{region 'Documentation'}
(*!
<summary>Neutral or held technical Error; task completion is reported separately.</summary>
*)
{endregion}
{attribute 'monitoring' := 'call'}
PROPERTY Result : E_Result //! Neutral or held technical Error; task completion is reported separately.
GET // PUBLIC
END_GET
END_PROPERTY

END_INTERFACE

// ---- Framework/Common/Interfaces/I_ResultAggregator.TcIO
{region 'Documentation'}
(*!
<summary>Contribution-only view of an owner-held result collection. Reset and result/counter access remain with the owner.</summary>
<description>
The owner resets and reads its concrete collection; a contribution hook only adds each owned result once. Contributions are immediate, not subscriptions, and no provider reference is retained. The owner limits a collection to 65535 contributions. Total includes neutral and Abort outcomes as well as Passed, Failed and Error; logging severity is a separate domain.
</description>
*)
{endregion}
INTERFACE I_ResultAggregator

{region 'Documentation'}
(*!
<summary>Adds one provider result immediately; a null provider contributes one Error. No provider reference is retained.</summary>
*)
{endregion}
METHOD AddProvider
VAR_INPUT
    Provider : I_ResultProvider; //! Result provider read immediately; zero contributes Error. No reference is retained.
END_VAR
END_METHOD

{region 'Documentation'}
(*!
<summary>Counts one contribution and combines Error &gt; Abort &gt; Failed &gt; Passed &gt; NotEvaluated.</summary>
*)
{endregion}
METHOD AddResult
VAR_INPUT
    Result : E_Result; //! Evaluation result to count as one contribution; severity is Error > Abort > Failed > Passed > NotEvaluated.
END_VAR
END_METHOD

END_INTERFACE

// ---- Framework/Common/Interfaces/I_ResultProvider.TcIO
{region 'Documentation'}
(*!
<summary>Read-only identity and result view; queries do not advance or modify the provider.</summary>
*)
{endregion}
INTERFACE I_ResultProvider

{region 'Documentation'}
(*!
<summary>Hierarchical identity supplied by the owning initialization path.</summary>
*)
{endregion}
{attribute 'monitoring' := 'variable'}
PROPERTY Name : STRING(GVL_Constants.NameLength) //! Hierarchical identity supplied by the owning initialization path.
GET // PUBLIC
END_GET
END_PROPERTY

{region 'Documentation'}
(*!
<summary>Current result by value; reading has no processing side effects.</summary>
*)
{endregion}
{attribute 'monitoring' := 'call'}
PROPERTY Result : E_Result //! Current result by value; reading has no processing side effects.
GET // PUBLIC
END_GET
END_PROPERTY

END_INTERFACE

// ---- Framework/EventBuffer/Interfaces/I_EventBuffer.TcIO
{region 'Documentation'}
(*!
<summary>Event storage initialization, administration, and value snapshots.</summary>
<description>
Bind one-based event storage and producer-owned status fields before administration. Keep them alive and stable and reinitialize after online change. The default service is single-task. Exactly one logical consumer acknowledges an epoch. External command handling and hierarchical reservation release belong to Run Control rather than this interface.
</description>
*)
{endregion}
INTERFACE I_EventBuffer

{region 'Documentation'}
(*!
<summary>Value snapshot of readable-range metadata.</summary>
*)
{endregion}
{attribute 'monitoring' := 'variable'}
PROPERTY FifoStatus : ST_FifoStatus //! Value snapshot of readable-range metadata.
GET // PUBLIC
END_GET
END_PROPERTY

{region 'Documentation'}
(*!
<summary>Bind one-based event storage and its producer-owned status fields for the service lifetime.</summary>
<description>
Establish an empty epoch; update the status fields internally after storage operations.

The default service requires lower bound 1 and physical length 3..32767; one ring position remains unused. Successful initialization clears the payload and begins a new empty epoch. Initialize owner reservation ledgers consistently; isolated reinitialization during execution is unsupported.
</description>
*)
{endregion}
METHOD Initialize : BOOL //! TRUE when storage is bound and usable; FALSE leaves the service uninitialized.
VAR_IN_OUT
    Buffer : ARRAY[*] OF ST_Event; //! Caller-owned event array, bound by address until reinitialization; keep storage alive and unchanged.
    FifoControl : ST_FifoStatus; //! Caller-owned FIFO status storage, retained and updated after buffer operations; must outlive the service.
    Status : ST_EventBufferStatus; //! Caller-owned event-sequence/loss snapshot, retained and updated by the service; must outlive it.
END_VAR
END_METHOD

{region 'Documentation'}
(*!
<summary>Release through the captured watermark; clear the caller&#x27;s field only if unchanged.</summary>
<description>
Use a current-epoch contiguous watermark after processing all preceding unread events. Zero is a no-op. Rejection or partial progress can still clear an unchanged request; inspect the actual DeletedSequenceId rather than treating command clearing as successful acknowledgement.
</description>
*)
{endregion}
METHOD ProcessDeleteRequest
VAR_IN_OUT
    SequenceId : UDINT; //! Inclusive deletion watermark; zero means no request. Cleared only if unchanged after processing.
END_VAR
END_METHOD

{region 'Documentation'}
(*!
<summary>Clear storage and epoch state while retaining a valid initialized binding.</summary>
<description>
A valid binding is required. The default service clears event storage, FIFO state, sequence, deletion watermark, loss count and aggregate reservations, retaining the binding. Owner-local accounting and external commands are handled by the Run Control integration path; they are not repaired here. Old-epoch acknowledgements become invalid.
</description>
*)
{endregion}
METHOD Reset
END_METHOD

{region 'Documentation'}
(*!
<summary>Value snapshot of sequence, deletion and loss status.</summary>
*)
{endregion}
{attribute 'monitoring' := 'variable'}
PROPERTY Status : ST_EventBufferStatus //! Value snapshot of sequence, deletion and loss status.
GET // PUBLIC
END_GET
END_PROPERTY

END_INTERFACE

// ---- Framework/EventBuffer/Interfaces/I_EventPublisher.TcIO
{region 'Documentation'}
(*!
<summary>PLC-side event publication and capacity view.</summary>
<description>
The default service is single-task and must be initialized with valid, stable storage before use. Publication copies the payload and assigns sequence/time; it does not consume an owner's reservation. Reservations are admission accounting, not storage or per-publication protection. Keep owner contributions consistent with the aggregate count and release them through their owner operations. Sequence exhaustion within an epoch is unsupported.
</description>
*)
{endregion}
INTERFACE I_EventPublisher

{region 'Documentation'}
(*!
<summary>Usable event positions, independent of occupancy and reservations; zero when invalid.</summary>
*)
{endregion}
{attribute 'monitoring' := 'call'}
PROPERTY Capacity : UINT //! Usable event positions, independent of occupancy and reservations; zero when invalid.
GET // PUBLIC
END_GET
END_PROPERTY

{region 'Documentation'}
(*!
<summary>Usable free event positions before reservations; zero when invalid.</summary>
*)
{endregion}
{attribute 'monitoring' := 'call'}
PROPERTY FreeEntryCount : UINT //! Usable free event positions before reservations; zero when invalid.
GET // PUBLIC
END_GET
END_PROPERTY

{region 'Documentation'}
(*!
<summary>Release only reservations, never events; FALSE changes neither count.</summary>
<description>
Requires an initialized valid binding, but no free capacity or valid FIFO indices.

The default service validates configuration and accounting even for a zero release. Free capacity and valid FIFO indices are not required. Destructive buffer reset clears the aggregate ledger, not stale owner-local contributions; use the coordinated owner release/reset path.
</description>
*)
{endregion}
METHOD FreeReservedSpace : BOOL //! TRUE after updating both reservation counts; FALSE leaves both unchanged.
VAR_INPUT
    EntryCount : UINT; //! Number of this owner's reserved entries to release; does not delete events.
END_VAR
VAR_IN_OUT
    OwnerReservedEntryCount : UINT; //! Owner's live reservation ledger; updated with the global count only on success, unchanged on rejection.
END_VAR
END_METHOD

{region 'Documentation'}
(*!
<summary>FIFO binding, configuration and indices are valid.</summary>
*)
{endregion}
{attribute 'monitoring' := 'call'}
PROPERTY IsValid : BOOL //! FIFO binding, configuration and indices are valid.
GET // PUBLIC
END_GET
END_PROPERTY

{region 'Documentation'}
(*!
<summary>Lost event count for producer diagnostics and aggregation.</summary>
*)
{endregion}
{attribute 'monitoring' := 'call'}
PROPERTY LostEventCount : UINT //! Lost event count for producer diagnostics and aggregation.
GET // PUBLIC
END_GET
END_PROPERTY

{region 'Documentation'}
(*!
<summary>Publish a value copy with producer-assigned SequenceId and UTC Timestamp.</summary>
<description>
Positive slot on success, zero when full, negative E_EventPublishResult on error.

The return describes the requested event. The default service may also attempt a capacity diagnostic after a successful insertion. That attempt can consume capacity or increase LostEventCount without changing the primary return. Publishing does not decrement an owner's reservation. Sequence numbers may be assigned before insertion succeeds; a nonzero loss count means an incomplete log.
</description>
*)
{endregion}
METHOD PublishEvent : INT //! Positive physical slot on success, zero when full, negative E_EventPublishResult on error.
VAR_INPUT
    Event : ST_Event; //! Event payload copied into the buffer; SequenceId and Timestamp are assigned by the publisher.
END_VAR
END_METHOD

{region 'Documentation'}
(*!
<summary>Aggregate producer reservations; not published externally.</summary>
*)
{endregion}
{attribute 'monitoring' := 'call'}
PROPERTY ReservedEntryCount : UINT //! Aggregate producer reservations; not published externally.
GET // PUBLIC
END_GET
END_PROPERTY

{region 'Documentation'}
(*!
<summary>Reserve additional event positions plus shared headroom; FALSE changes neither count.</summary>
<description>
Requires valid initialized configuration and a consistent owner contribution; positive requests also require valid indices.

For the default service, positive requests require free capacity for the updated aggregate count plus shared headroom. A zero request checks configuration and owner contribution but bypasses index and capacity checks. Both ledgers change together on success; no event is created. Keep the owner ledger unchanged by unrelated code.
</description>
*)
{endregion}
METHOD ReserveSpace : BOOL //! TRUE after updating both reservation counts; FALSE leaves both unchanged.
VAR_INPUT
    EntryCount : UINT; //! Additional number of event entries to reserve for this owner.
    HeadroomEntryCount : UINT; //! Shared free entries checked for positive requests; not added to the owner's reservation.
END_VAR
VAR_IN_OUT
    OwnerReservedEntryCount : UINT; //! Owner's live reservation ledger; updated with the global count only on success, unchanged on rejection.
END_VAR
END_METHOD

END_INTERFACE

// ---- Framework/Preparation/Interfaces/I_Preparation.TcIO
{region 'Documentation'}
(*!
<summary>Read-only Preparation view; querying does not execute resource actions.</summary>
<description>
This interface exposes only the last reported Status by value. The owner calls the concrete Preparation cyclically with Enable and its resource-specific bindings; the interface provides no generic activation, initialization or reset operation.
</description>
*)
{endregion}
INTERFACE I_Preparation

{region 'Documentation'}
(*!
<summary>Current Preparation status by value; querying does not execute resource actions.</summary>
*)
{endregion}
PROPERTY Status : ST_PreparationStatus //! Current Preparation status by value; querying does not execute resource actions.
GET // PUBLIC
END_GET
END_PROPERTY

END_INTERFACE

// ---- Framework/RunControl/Interfaces/I_RunControl.TcIO
{region 'Documentation'}
(*!
<summary>Run Control request and status view; the execution owner calls the concrete FB cyclically.</summary>
<description>
Request methods record same-task intent; they do not execute the lifecycle synchronously. Repeated requests coalesce and regular processing applies Reset over Abort over Start. Status is a stored value snapshot. Name and Result are inherited from I_ResultProvider. The concrete owner must still be called cyclically, including after completion.
</description>
*)
{endregion}
INTERFACE I_RunControl EXTENDS I_ResultProvider

{region 'Documentation'}
(*!
<summary>Records an abort request for regular lifecycle processing.</summary>
*)
{endregion}
METHOD RequestAbort
END_METHOD

{region 'Documentation'}
(*!
<summary>Records a reset request for regular lifecycle processing.</summary>
*)
{endregion}
METHOD RequestReset
END_METHOD

{region 'Documentation'}
(*!
<summary>Records a start request for regular lifecycle processing.</summary>
*)
{endregion}
METHOD RequestStart
END_METHOD

{region 'Documentation'}
(*!
<summary>Current owner status snapshot; reading does not execute lifecycle processing.</summary>
*)
{endregion}
PROPERTY Status : ST_RunControlStatus //! Current owner status snapshot; reading does not execute lifecycle processing.
GET // PUBLIC
END_GET
END_PROPERTY

END_INTERFACE

// ---- Framework/TestCases/Interfaces/I_TestCase.TcIO
{region 'Documentation'}
(*!
<summary>Typed owner status with the shared child orchestration view.</summary>
<description>
Adds only the typed Status snapshot to I_Orchestratable. Lifecycle requests, readiness/state, initialization, reservation operations, execution slot and inherited identity/result belong to that shared child view. Requests do not execute the concrete FB. The owning Suite calls the concrete instance cyclically; status reads do not refresh it.
</description>
*)
{endregion}
INTERFACE I_TestCase EXTENDS I_Orchestratable

{region 'Documentation'}
(*!
<summary>Return the latest typed Test Case status by value without executing lifecycle, Preparation or Assertion work.</summary>
*)
{endregion}
PROPERTY Status : ST_TestCaseStatus //! Return the latest typed Test Case status by value without executing lifecycle, Preparation or Assertion work.
GET // PUBLIC
END_GET
END_PROPERTY

END_INTERFACE

// ---- Framework/TestSuites/Interfaces/I_TestSuite.TcIO
{region 'Documentation'}
(*!
<summary>Typed owner status with the shared child orchestration view.</summary>
<description>
Adds only typed Status to I_Orchestratable; shared requests, readiness/state, initialization, reservation operations, slot and inherited identity/result remain in that view. The owner invokes the concrete FB cyclically; interface requests and getters do not execute it. Production composition and the explicitly childless mock have different internal responsibilities.
</description>
*)
{endregion}
INTERFACE I_TestSuite EXTENDS I_Orchestratable

{region 'Documentation'}
(*!
<summary>Current owner status snapshot; reading does not execute lifecycle processing.</summary>
*)
{endregion}
PROPERTY Status : ST_TestSuiteStatus //! Current owner status snapshot; reading does not execute lifecycle processing.
GET // PUBLIC
END_GET
END_PROPERTY

END_INTERFACE

// ---- Runtime/MAIN.TcPOU
{region 'Documentation'}
(*!
<summary>Initializes the selftest hierarchy on the first task cycle and executes its command adapter and root.</summary>
<description>
Assign MAIN once to the single cyclic task that owns the hierarchy. A nonpositive current task
index skips all work. On FirstCycle, clear old commands through the adapter, initialize the
actual Event Stream storage/status, then initialize the SelfTests root with that same buffer service.
The library's default publisher must refer to the matching service before configuration diagnostics.

Normal processing calls the command adapter before the concrete root on every valid task call,
including after initialization failure or lifecycle completion. The stored initialization outcomes
are diagnostic values, not cyclic execution gates; failed owner setup prevents normal child work
inside the base. There is no automatic cyclic initialization retry or automatic Start of tests.

Successful root initialization queues its initial lifecycle Reset; readiness is established over
subsequent cycles. Rebuilding setup requires configuration reactivation or PLC Cold Reset and the
coordinated first-cycle path. Normal Stop/Start and lifecycle Reset do not rebuild configuration.
This executable selftest composition is outside the packaged library and consumer API reference.
</description>
*)
{endregion}
PROGRAM MAIN
VAR
    {attribute 'TcNoSymbol'}
    FRunControl : RunControl; //! Statically owned selftest root; invoked once after command intake on every valid task call.
    {attribute 'TcNoSymbol'}
    FCommandAdapter : RunControlCommandAdapter; //! Owner-local command sampler; initialized before the Event Buffer and called before the root.
    {attribute 'TcNoSymbol'}
    FEventBufferInitialized : BOOL; //! Last first-cycle Event Buffer initialization outcome; diagnostic only, not a cyclic call gate.
    {attribute 'TcNoSymbol'}
    FFrameworkInitialized : BOOL; //! Last first-cycle hierarchy initialization outcome; TRUE does not yet imply Idle or Ready.
END_VAR
VAR_TEMP
    TaskIndex : DINT; //! Current cyclic PLC task index; nonpositive values skip initialization and execution.
END_VAR

TaskIndex := Tc2_System.GETCURTASKINDEXEX();
IF TaskIndex <= 0 THEN
    RETURN;
END_IF;

IF TwinCAT_SystemInfoVarList._TaskInfo[TaskIndex].FirstCycle THEN
    FCommandAdapter.Initialize(ControlData := GVL_UnitTest.RunControl.ControlData);

    FEventBufferInitialized := GVL_EventBuffer.Instance.Initialize(Buffer := GVL_UnitTest.EventStream.Buffer,
        FifoControl := GVL_UnitTest.EventStream.FifoControl,
        Status := GVL_UnitTest.EventStream.Status);

    FFrameworkInitialized := FRunControl.Initialize(Name := 'SelfTests',
        EventBuffer := GVL_EventBuffer.Instance);
END_IF;

FCommandAdapter(RunControl := FRunControl,
    Commands := GVL_UnitTest.RunControl.ControlData.Cmd);
FRunControl(ControlData := GVL_UnitTest.RunControl.ControlData);

END_PROGRAM

// ---- SelfTests/RunControl/RunControl.TcPOU
{region 'Documentation'}
(*!
<summary>Composes the selftest Suites and forwards the external communication storage to the root base.</summary>
*)
{endregion}
FUNCTION_BLOCK RunControl EXTENDS RunControlBase
VAR
    FSmoke : TestSuite_Smoke;
    FPreparation : TestSuite_Preparation;
    FTestCaseLifecycle : TestSuite_TestCaseLifecycle;
    FOrchestratorTests : TestSuite_Orchestrator;
    FSerialOrchestration : TestSuite_SerialOrchestration;
    FParallelOrchestration : TestSuite_ParallelOrchestration;
    FParallelSlotsOrchestration : TestSuite_ParallelSlotsOrchestration;
    FSuiteBuilderTests : TestSuite_TestSuiteConfigurationBuilder;
    FRunControlBuilderTests : TestSuite_RunControlConfigurationBuilder;
    FTestSuites : ARRAY[1..SuiteCapacity] OF I_TestSuite;
    FTestSuiteLifecycle : TestSuite_TestSuiteLifecycle;
    FRunControlLifecycle : TestSuite_RunControlLifecycle;
    FCommandAdapter : TestSuite_CommandAdapter;
    FEventDelivery : TestSuite_EventDelivery;
    FEventReservation : TestSuite_EventReservation;
    FEventBufferReset : TestSuite_EventBufferReset;
    FAssertionLifecycle : TestSuite_AssertionLifecycle;
    FAssertionComparisons : TestSuite_AssertionComparisons;
    FAssertionFloatingPoint : TestSuite_AssertionFloatingPoint;
    FAssertionObservation : TestSuite_AssertionObservation;
    FAssertionText : TestSuite_AssertionText;
    FAssertionArrays : TestSuite_AssertionArrays;
    FAssertionVariants : TestSuite_AssertionVariants;
END_VAR
VAR CONSTANT
    SuiteCapacity : UINT := 22;
END_VAR

SUPER^(ControlData := ControlData);

{region 'Documentation'}
(*!
<summary>Initializes and registers the selftest Suites serially. Root and Suite Reset timeouts allow 15 seconds for event-consumer backpressure.</summary>
*)
{endregion}
METHOD PROTECTED Configure
VAR_IN_OUT
    // SA0167: Borrowed builder; VAR_IN_OUT creates no temporary instance.
    {attribute 'analysis' := '-167'}
    Builder : RunControlConfigurationBuilder; //! Borrowed owner configuration builder used only during this Configure call; register this owner's concrete children.
END_VAR
VAR
    SuiteConfig : ST_TestSuiteConfig;
END_VAR
FConfig.Timeout := T#60s;
FConfig.ResetTimeout := T#15s;
SuiteConfig.ResetTimeout := T#15s;

Builder.Initialize(Mode := E_OrchestrationMode.Serial,
    TestSuites := FTestSuites);

FSmoke.Initialize(Parent := THIS^,
    SuiteName := 'Smoke',
    Config := SuiteConfig);
Builder.Register(TestSuite := FSmoke);

FPreparation.Initialize(Parent := THIS^,
    SuiteName := 'Preparation',
    Config := SuiteConfig);
Builder.Register(TestSuite := FPreparation);

FTestCaseLifecycle.Initialize(Parent := THIS^,
    SuiteName := 'TestCaseLifecycle',
    Config := SuiteConfig);
Builder.Register(TestSuite := FTestCaseLifecycle);

FOrchestratorTests.Initialize(Parent := THIS^,
    SuiteName := 'Orchestrator',
    Config := SuiteConfig);
Builder.Register(TestSuite := FOrchestratorTests);

FSerialOrchestration.Initialize(Parent := THIS^,
    SuiteName := 'SerialOrchestration',
    Config := SuiteConfig);
Builder.Register(TestSuite := FSerialOrchestration);

FParallelOrchestration.Initialize(Parent := THIS^,
    SuiteName := 'ParallelOrchestration',
    Config := SuiteConfig);
Builder.Register(TestSuite := FParallelOrchestration);

FParallelSlotsOrchestration.Initialize(Parent := THIS^,
    SuiteName := 'ParallelSlotsOrchestration',
    Config := SuiteConfig);
Builder.Register(TestSuite := FParallelSlotsOrchestration);

FSuiteBuilderTests.Initialize(Parent := THIS^,
    SuiteName := 'SuiteBuilder',
    Config := SuiteConfig);
Builder.Register(TestSuite := FSuiteBuilderTests);

FRunControlBuilderTests.Initialize(Parent := THIS^,
    SuiteName := 'RunControlBuilder',
    Config := SuiteConfig);
Builder.Register(TestSuite := FRunControlBuilderTests);

FTestSuiteLifecycle.BindSubjectParent(Parent := THIS^);
FTestSuiteLifecycle.Initialize(Parent := THIS^,
    SuiteName := 'TestSuiteLifecycle',
    Config := SuiteConfig);
Builder.Register(TestSuite := FTestSuiteLifecycle);

FRunControlLifecycle.Initialize(Parent := THIS^,
    SuiteName := 'RunControlLifecycle',
    Config := SuiteConfig);
Builder.Register(TestSuite := FRunControlLifecycle);

FCommandAdapter.Initialize(Parent := THIS^,
    SuiteName := 'CommandAdapter',
    Config := SuiteConfig);
Builder.Register(TestSuite := FCommandAdapter);

FEventDelivery.Initialize(Parent := THIS^,
    SuiteName := 'EventDelivery',
    Config := SuiteConfig);
Builder.Register(TestSuite := FEventDelivery);

FEventReservation.BindSubjectParent(Parent := THIS^);
FEventReservation.Initialize(Parent := THIS^,
    SuiteName := 'EventReservation',
    Config := SuiteConfig);
Builder.Register(TestSuite := FEventReservation);

FEventBufferReset.Initialize(Parent := THIS^,
    SuiteName := 'EventBufferReset',
    Config := SuiteConfig);
Builder.Register(TestSuite := FEventBufferReset);

FAssertionLifecycle.Initialize(Parent := THIS^,
    SuiteName := 'AssertionLifecycle',
    Config := SuiteConfig);
Builder.Register(TestSuite := FAssertionLifecycle);

FAssertionComparisons.Initialize(Parent := THIS^,
    SuiteName := 'AssertionComparisons',
    Config := SuiteConfig);
Builder.Register(TestSuite := FAssertionComparisons);

FAssertionFloatingPoint.Initialize(Parent := THIS^,
    SuiteName := 'AssertionFloatingPoint',
    Config := SuiteConfig);
Builder.Register(TestSuite := FAssertionFloatingPoint);

FAssertionObservation.Initialize(Parent := THIS^,
    SuiteName := 'AssertionObservation',
    Config := SuiteConfig);
Builder.Register(TestSuite := FAssertionObservation);

FAssertionText.Initialize(Parent := THIS^,
    SuiteName := 'AssertionText',
    Config := SuiteConfig);
Builder.Register(TestSuite := FAssertionText);

FAssertionArrays.Initialize(Parent := THIS^,
    SuiteName := 'AssertionArrays',
    Config := SuiteConfig);
Builder.Register(TestSuite := FAssertionArrays);

FAssertionVariants.Initialize(Parent := THIS^,
    SuiteName := 'AssertionVariants',
    Config := SuiteConfig);
Builder.Register(TestSuite := FAssertionVariants);
END_METHOD

{region 'Documentation'}
(*!
<summary>Returns the registered Suite from the same array used during configuration.</summary>
*)
{endregion}
METHOD PUBLIC GetTestSuite : I_TestSuite //! Typed Suite interface at the original array index; zero when no entry is available.
VAR_INPUT
    Index : DINT; //! Original occupied child-array index, rather than an ordinal position.
END_VAR
GetTestSuite := 0;
IF (ChildCount = 0) OR (Index < ChildArrayLowerBound)
    OR (DINT_TO_LINT(Index) >= DINT_TO_LINT(ChildArrayLowerBound) + UINT_TO_LINT(ChildCount)) THEN
    RETURN;
END_IF;

GetTestSuite := FTestSuites[Index];
END_METHOD

{region 'Documentation'}
(*!
<summary>Calls each owned Suite once per initialized root cycle, including completion.</summary>
*)
{endregion}
METHOD PROTECTED ProcessTestSuites
FSmoke();
FPreparation();
FTestCaseLifecycle();
FOrchestratorTests();
FSerialOrchestration();
FParallelOrchestration();
FParallelSlotsOrchestration();
FSuiteBuilderTests();
FRunControlBuilderTests();

FTestSuiteLifecycle();
FRunControlLifecycle();

FCommandAdapter();

FEventDelivery();

FEventReservation();
FEventBufferReset();
FAssertionLifecycle();
FAssertionComparisons();
FAssertionFloatingPoint();
FAssertionObservation();

FAssertionText();

FAssertionArrays();
FAssertionVariants();
END_METHOD

END_FUNCTION_BLOCK

// ---- Framework/RunControl/POU/RunControlBase.TcPOU
{region 'Documentation'}
(*!
<summary>Root lifecycle and orchestration of the application's static Suite collection.</summary>
<description>
The PLC program initializes the Event Buffer and publisher before Initialize. Implement
Configure, GetTestSuite and ProcessTestSuites; forward ControlData to SUPER^() once per task
cycle.

Run the external command adapter before this FB. Buffer commands are handled first; only Name
and Status are projected after lifecycle processing. CompletionDelay belongs to this root, not to
its Orchestrator.

Continue cyclic calls after Completed so descendants can finish outstanding work and status
can refresh. This does not reopen the finalized root result.

In Completing, Result and Aggregation are published once before CompletionDelay elapses. The
final transition occurs on a later call even for zero delay. Invalid delay timing emits a diagnostic
and completes without changing published results.
</description>
*)
{endregion}
FUNCTION_BLOCK ABSTRACT RunControlBase IMPLEMENTS I_RunControl, I_OrchestratableCollection
VAR_IN_OUT
    ControlData : ST_RunControl; //! External communication storage; BufferCmd is processed first, Name and Status are projected last.
END_VAR
VAR
    /// Instance binding; derived test adapters may assign it before first use.
    FEventPublisher : I_EventPublisher;
    FName : STRING(GVL_Constants.NameLength);
    FResourceName : STRING(GVL_Constants.ResourceNameLength);
    FConfig : ST_RunConfig;
    FEventBuffer : I_EventBuffer;
    FCollectionConfiguration : ST_TestSuiteCollectionConfig;
    FOrchestrator : I_Orchestrator;
    FDefaultOrchestrator : Orchestrator;
    FInitialized : BOOL;
    FHasTimeout : BOOL;
    FHasResetTimeout : BOOL;
    FHasAbortTimeout : BOOL;
    FCheckingInitialization : BOOL;
    FConfigError : BOOL;
    FStatus : ST_RunControlStatus;
    FResult : E_Result := E_Result.NotEvaluated;
    FState : E_State := E_State.Uninitialized;
    FMethodRequests : ST_Command;
    FExecutionTimer : Stopwatch;
    FStateTimer : Stopwatch;
    FAggregator : ResultAggregator;
    FTestSuiteCountInactive : UINT;
    FTestSuiteCountIdle : UINT;
    FTestSuiteCountRunning : UINT;
    FTestSuiteCountCompleted : UINT;
    FTestSuiteCountError : UINT;
    FCollectionValid : BOOL;
    FChildrenError : BOOL;
    FChildrenAborted : BOOL;
    FChildrenCompleted : BOOL;
    FChildrenAbortFinished : BOOL;
    FFinalizationPublished : BOOL;
END_VAR
VAR_TEMP
    Requests : ST_Command;
    OrchestratorTask : E_OrchestratorTask;
END_VAR

ProcessBufferCommands(Commands := ControlData.BufferCmd);
ProcessRequests(InputRequests := FMethodRequests, Requests => Requests);

FExecutionTimer.Update();
FStateTimer.Update();

Sequencer(Requests := Requests);

IF IsInitialized THEN
    OrchestratorTask := MapOrchestratorTask(State := FState,
        CurrentTask := FOrchestrator.CurrentTask);
    FOrchestrator.Execute(Task := OrchestratorTask);

    ProcessTestSuites();
    AggregateResults();
END_IF;

UpdateResult();
UpdateStatus();
EmitFinalizationEvents();

ControlData.Name := FName;
ControlData.Status := FStatus;

{region 'Documentation'}
(*!
<summary>Aggregates results and execution counters after child calls; refreshes observations from the same snapshots.</summary>
*)
{endregion}
METHOD PRIVATE AggregateResults
VAR
    Count : UINT;
    FirstIndex : DINT;
    LastIndex : DINT;
    Index : LINT;
    ChildStatus : ST_TestSuiteStatus;
    ChildResult : E_Result;
END_VAR
Count := ChildCount;
FTestSuiteCountInactive := 0;
FTestSuiteCountIdle := 0;
FTestSuiteCountRunning := 0;
FTestSuiteCountCompleted := 0;
FTestSuiteCountError := 0;
FAggregator.Reset();
FCollectionValid := FALSE;
FChildrenCompleted := FALSE;
FChildrenAbortFinished := FALSE;
FChildrenError := FALSE;
FChildrenAborted := FALSE;

IF NOT FInitialized OR (Count = 0) THEN
    RETURN;
END_IF;
FirstIndex := ChildArrayLowerBound;
LastIndex := ChildArrayUpperBound;
IF DINT_TO_LINT(LastIndex) - DINT_TO_LINT(FirstIndex) + 1 < UINT_TO_LINT(Count) THEN
    RETURN;
END_IF;

FCollectionValid := TRUE;
FChildrenCompleted := TRUE;
FChildrenAbortFinished := TRUE;
FOR Index := DINT_TO_LINT(FirstIndex) TO DINT_TO_LINT(FirstIndex) + UINT_TO_LINT(Count) - 1 DO
    IF NOT ObserveTestSuite(Child := GetTestSuite(Index := LINT_TO_DINT(Index)),
        ChildStatus => ChildStatus) THEN
        FTestSuiteCountError := FTestSuiteCountError + 1;
        FAggregator.AddResult(Result := E_Result.Error);
        CONTINUE;
    END_IF;

    ChildResult := ChildStatus.Execution.Result;
    CASE ChildResult OF
        E_Result.NotEvaluated, E_Result.Passed, E_Result.Failed, E_Result.Abort, E_Result.Error:
            FAggregator.AddResult(Result := ChildResult);
    ELSE
        ChildResult := E_Result.Error;
        FAggregator.AddResult(Result := ChildResult);
    END_CASE;

    CASE ChildStatus.Execution.ExecutionStatus OF
        E_ExecutionStatus.Inactive:
            FTestSuiteCountInactive := FTestSuiteCountInactive + 1;
        E_ExecutionStatus.Idle:
            FTestSuiteCountIdle := FTestSuiteCountIdle + 1;
        E_ExecutionStatus.Running:
            FTestSuiteCountRunning := FTestSuiteCountRunning + 1;
        E_ExecutionStatus.Completed:
            FTestSuiteCountCompleted := FTestSuiteCountCompleted + 1;
    ELSE
        // Transitional execution states have no dedicated counter in the status contract.
    END_CASE;
    IF (ChildStatus.Execution.ExecutionStatus = E_ExecutionStatus.Error) OR (ChildResult = E_Result.Error) THEN
        FTestSuiteCountError := FTestSuiteCountError + 1;
    END_IF;

END_FOR;
END_METHOD

{region 'Documentation'}
(*!
<summary>Applies permitted owner transitions; rejects others with state-dependent diagnostics and Error escalation while leaving FState unchanged.</summary>
*)
{endregion}
METHOD PRIVATE ChangeState
VAR_INPUT
    NewState : E_State; //! Requested owner lifecycle destination; identical state is a no-op and rejected transitions do not change FState.
END_VAR
IF NewState = FState THEN
    RETURN;
END_IF;
IF NOT IsStateTransitionAllowed(NewState := NewState) THEN
    CASE FState OF
        E_State.Uninitialized:
            RETURN;

        E_State.Completing, E_State.Completed:
            PublishEvent(Event := CreateInvalidStateTransitionEvent(OwnerScope := E_OwnerScope.RunControl,
                Name := FName,
                ResourceName := FResourceName,
                StateOld := FState,
                StateNew := NewState));
    ELSE
        IF FResult <> E_Result.Error THEN
            PublishEvent(Event := CreateInvalidStateTransitionEvent(OwnerScope := E_OwnerScope.RunControl,
                Name := FName,
                ResourceName := FResourceName,
                StateOld := FState,
                StateNew := NewState));
        END_IF;
        FResult := E_Result.Error;
    END_CASE;
    RETURN;
END_IF;

CASE NewState OF
    E_State.Uninitialized:
        FExecutionTimer.Reset();
        FStateTimer.Start();
        FResult := E_Result.NotEvaluated;
    E_State.Reset:
        FHasTimeout := FALSE;
        FHasResetTimeout := FALSE;
        FHasAbortTimeout := FALSE;
        FFinalizationPublished := FALSE;
        FAggregator.Reset();
        IF (FState = E_State.Starting) OR (FState = E_State.Running) OR (FState = E_State.Completing)
            OR (FState = E_State.Aborting) OR (FState = E_State.AbortingFromError) THEN
            PublishEvent(Event := CreateResetWarningEvent(OwnerScope := E_OwnerScope.RunControl,
                Name := FName,
                ResourceName := FResourceName,
                State := FState));
        END_IF;
        FExecutionTimer.Reset();
        FStateTimer.Start();
        FResult := E_Result.NotEvaluated;
    E_State.Idle:
        FStateTimer.Start();
    E_State.Starting:
        FStateTimer.Start();
        FExecutionTimer.Start();
    E_State.Running:
        FStateTimer.Start();
    E_State.Completing:
        FExecutionTimer.Stop();
        FStateTimer.Start();
    E_State.Completed:
        FStateTimer.Start();
    E_State.Aborting:
        FExecutionTimer.Stop();
        FStateTimer.Start();
        IF FResult <> E_Result.Error THEN
            FResult := E_Result.Abort;
        END_IF;
    E_State.AbortingFromError:
        FExecutionTimer.Stop();
        IF FState <> E_State.Aborting THEN
            FStateTimer.Start();
        END_IF;
        FResult := E_Result.Error;
ELSE
    RETURN;
END_CASE;
PublishEvent(Event := CreateStateTransitionEvent(OwnerScope := E_OwnerScope.RunControl,
    Name := FName,
    ResourceName := FResourceName,
    StateOld := FState,
    StateNew := NewState));
FState := NewState;
END_METHOD

{region 'Documentation'}
(*!
<summary>Validates timeouts, the initialized Orchestrator and every registered child.</summary>
<description>
Called after builder finalization and helper initialization. An override must include
SUPER^.CheckInitialization(), preserve failure and check any additional application setup.

Timeout, ResetTimeout and AbortTimeout must be positive. CompletionDelay may be zero. The base
reports its first failed check; FALSE prevents successful initialization.
</description>
*)
{endregion}
METHOD PROTECTED CheckInitialization : BOOL //! TRUE when the configured setup is valid; FALSE reports invalid setup and prevents initialization.
VAR
    Index : LINT;
    Child : I_TestSuite;
END_VAR
CheckInitialization := FALSE;
IF (FConfig.Timeout = T#0ms) OR (FConfig.ResetTimeout = T#0ms) OR (FConfig.AbortTimeout = T#0ms) THEN
    PublishInitializationError(Message := 'Run timeouts must be greater than zero.');
    RETURN;
END_IF;
IF NOT FOrchestrator.IsInitialized THEN
    PublishInitializationError(Message := 'Orchestrator initialization is invalid.');
    RETURN;
END_IF;
IF (ChildCount = 0)
    OR (DINT_TO_LINT(ChildArrayUpperBound) - DINT_TO_LINT(ChildArrayLowerBound) + 1 < UINT_TO_LINT(ChildCount)) THEN
    PublishInitializationError(Message := 'Invalid registered Test Suite range.');
    RETURN;
END_IF;
FOR Index := DINT_TO_LINT(ChildArrayLowerBound) TO DINT_TO_LINT(ChildArrayLowerBound) + UINT_TO_LINT(ChildCount) - 1 DO
    Child := GetTestSuite(Index := LINT_TO_DINT(Index));
    IF Child = 0 THEN
        PublishInitializationError(Message := CONCAT('Missing Test Suite at index ', LINT_TO_STRING(Index)));
        RETURN;
    END_IF;
    IF NOT Child.IsInitialized THEN
        PublishInitializationError(Message := CONCAT('Test Suite is not initialized: ', Child.Name));
        RETURN;
    END_IF;
END_FOR;
CheckInitialization := TRUE;
END_METHOD

{region 'Documentation'}
(*!
<summary>Actual lower array bound; zero when collection metadata is unavailable.</summary>
*)
{endregion}
{attribute 'monitoring' := 'call'}
PROPERTY PUBLIC ChildArrayLowerBound : DINT //! Actual lower array bound; zero when collection metadata is unavailable.
GET // PUBLIC
ChildArrayLowerBound := 0;
IF NOT (FInitialized OR FCheckingInitialization) OR NOT FCollectionConfiguration.IsValid THEN
    RETURN;
END_IF;
ChildArrayLowerBound := FCollectionConfiguration.FirstIndex;
END_GET
END_PROPERTY

{region 'Documentation'}
(*!
<summary>Actual upper array bound including unused capacity; zero when unavailable.</summary>
*)
{endregion}
{attribute 'monitoring' := 'call'}
PROPERTY PUBLIC ChildArrayUpperBound : DINT //! Actual upper array bound including unused capacity; zero when unavailable.
GET // PUBLIC
ChildArrayUpperBound := 0;
IF NOT (FInitialized OR FCheckingInitialization) OR NOT FCollectionConfiguration.IsValid THEN
    RETURN;
END_IF;
ChildArrayUpperBound := FCollectionConfiguration.LastIndex;
END_GET
END_PROPERTY

{region 'Documentation'}
(*!
<summary>Registered population; zero outside setup validation or successful
initialization.</summary>
*)
{endregion}
{attribute 'monitoring' := 'call'}
PROPERTY PUBLIC ChildCount : UINT //! Registered population; zero outside setup validation or successful initialization.
GET // PUBLIC
ChildCount := 0;
IF NOT (FInitialized OR FCheckingInitialization) OR NOT FCollectionConfiguration.IsValid THEN
    RETURN;
END_IF;
ChildCount := FCollectionConfiguration.Count;
END_GET
END_PROPERTY

{region 'Documentation'}
(*!
<summary>Initializes and registers this owner's static Suites.</summary>
<description>
Set FConfig and optional FResourceName. The owner identity is already established. Initialize
owned children, bind the local interface array through Builder.Initialize, select the mode, and use
Register or RegisterWithSlot as appropriate.

The base calls Finalize after this hook and retains only validated configuration values; it
then initializes the Orchestrator and calls CheckInitialization. Do not retain the borrowed
RunControlConfigurationBuilder or its temporary storage binding.

Implement GetTestSuite against that same array and keep the composition fixed until full
hierarchical reinitialization. This abstract hook has no base implementation to call.
</description>
*)
{endregion}
METHOD PROTECTED ABSTRACT Configure
VAR_IN_OUT
    // SA0167: Borrowed builder; VAR_IN_OUT creates no temporary instance.
    {attribute 'analysis' := '-167'}
    Builder : RunControlConfigurationBuilder; //! Borrowed setup builder; initialize and register children during Configure only. The base calls Finalize afterwards.
END_VAR
(* Builder.Initialize(Mode := E_OrchestrationMode.Serial,
    TestSuites := FTestSuites);
FExample.Initialize(Parent := THIS^,
    SuiteName := 'Example',
    Config := ExampleConfig);
Builder.Register(TestSuite := FExample);
Initialize and register each owned Suite; use RegisterWithSlot for ParallelSlots.
Keep the default FConfig values or assign the Run Control timing configuration here.
*)
END_METHOD

{region 'Documentation'}
(*!
<summary>Publishes Result then Aggregation once on entry to Completing; publication failure is not retried.</summary>
<description>
The final owner result and emitted payloads remain held; current status counters continue to refresh.
</description>
*)
{endregion}
METHOD PRIVATE EmitFinalizationEvents
VAR
    Message : STRING(GVL_Constants.MessageLength);
    LostEventCount : UINT;
END_VAR
IF (FState <> E_State.Completing) OR FFinalizationPublished THEN
    RETURN;
END_IF;

CASE FResult OF
    E_Result.Passed:
        Message := 'Run completed.';
    E_Result.Failed:
        Message := 'Run completed with failed result.';
    E_Result.Error:
        Message := 'Run completed with error.';
    E_Result.Abort:
        Message := 'Run aborted.';
ELSE
    Message := 'Run completed without evaluated result.';
END_CASE;

PublishEvent(Event := CreateResultEvent(OwnerScope := E_OwnerScope.RunControl,
    Name := FName,
    ResourceName := FResourceName,
    State := FState,
    Result := FResult,
    Message := Message));

LostEventCount := EventPublisher.LostEventCount;
PublishEvent(Event := CreateRunAggregationEvent(Name := FName,
    Status := FStatus,
    LostEventCount := LostEventCount));

FFinalizationPublished := TRUE;
END_METHOD

{region 'Documentation'}
(*!
<summary>Latches the technical Run Control error and emits its first diagnostic; does not change state.</summary>
*)
{endregion}
METHOD PRIVATE Error
VAR_INPUT
    Message : STRING(GVL_Constants.MessageLength); //! Framework diagnostic text emitted only when first escalating a mutable owner result to Error.
END_VAR
IF (FState = E_State.Uninitialized) OR (FState = E_State.Completed) OR FFinalizationPublished THEN
    RETURN;
END_IF;
IF FResult <> E_Result.Error THEN
    PublishEvent(Event := CreateFrameworkEvent(Name := FName,
        ResourceName := FResourceName,
        State := FState,
        Severity := E_EventSeverity.Error,
        Message := Message));
END_IF;
FResult := E_Result.Error;
END_METHOD

{region 'Documentation'}
(*!
<summary>Returns this instance's retained event-publication service.</summary>
<description>
If the local binding is zero, the getter takes GVL_EventBuffer.Publisher on access. An
established binding is retained; Initialize and lifecycle Reset do not replace it.

The default must be bound before first diagnostic use. Controlled test adapters may assign the
protected field before use. This getter performs no event publication, lifecycle processing or
reservation change.
</description>
*)
{endregion}
{attribute 'monitoring' := 'variable'}
PROPERTY PUBLIC EventPublisher : I_EventPublisher //! Returns this instance's retained event-publication service.
GET // PUBLIC
IF FEventPublisher = 0 THEN
    FEventPublisher := GVL_EventBuffer.Publisher;
END_IF;
EventPublisher := FEventPublisher;
END_GET
END_PROPERTY

{region 'Documentation'}
(*!
<summary>Returns the common view from the typed owner collection without executing the
child.</summary>
*)
{endregion}
METHOD PUBLIC FINAL GetChild : I_Orchestratable //! Registered child interface at Index; zero for an invalid or unoccupied index.
VAR_INPUT
    Index : DINT; //! Original child-array index, not a registration ordinal; valid children occupy LowerBound through LowerBound + Count - 1.
END_VAR
GetChild := 0;
IF (ChildCount = 0) OR (Index < ChildArrayLowerBound)
    OR (DINT_TO_LINT(Index) >= DINT_TO_LINT(ChildArrayLowerBound) + UINT_TO_LINT(ChildCount)) THEN
    RETURN;
END_IF;
GetChild := GetTestSuite(Index := Index);
END_METHOD

{region 'Documentation'}
(*!
<summary>Returns a registered child from the concrete owner's interface array.</summary>
<description>
Implement lookup in the same array configured by Configure, using its actual array index
rather than a hard-coded registration ordinal. Registration can reorder entries by slot.

Check the occupied range starting at ChildArrayLowerBound for ChildCount entries and return
zero outside it. Do not access unused capacity, execute the child, or cache a setup-time array
address. This abstract method has no base implementation.
</description>
*)
{endregion}
METHOD PUBLIC ABSTRACT GetTestSuite : I_TestSuite //! Registered child interface at Index; zero for an invalid or unoccupied index.
VAR_INPUT
    Index : DINT; //! Original child-array index, not a registration ordinal; valid children occupy LowerBound through LowerBound + Count - 1.
END_VAR
(* GetTestSuite := 0;
IF (ChildCount = 0) OR (Index < ChildArrayLowerBound)
    OR (DINT_TO_LINT(Index) >= DINT_TO_LINT(ChildArrayLowerBound) + UINT_TO_LINT(ChildCount)) THEN
    RETURN;
END_IF;
GetTestSuite := FTestSuites[Index];
*)
END_METHOD

{region 'Documentation'}
(*!
<summary>Reports a detected Abort timeout until Initialize or entry into a new Reset.</summary>
<description>
An expired abort deadline finishes through Completing with Error. Escalation from Aborting to
AbortingFromError does not restart that deadline.
</description>
*)
{endregion}
{attribute 'monitoring' := 'call'}
PROPERTY PUBLIC HasAbortTimeout : BOOL //! Reports a detected Abort timeout until Initialize or entry into a new Reset.
GET // PUBLIC
HasAbortTimeout := FHasAbortTimeout;
END_GET
END_PROPERTY

{region 'Documentation'}
(*!
<summary>Reports the current owner error condition used by status projection.</summary>
*)
{endregion}
{attribute 'monitoring' := 'call'}
PROPERTY PUBLIC HasError : BOOL //! Reports the current owner error condition used by status projection.
GET // PUBLIC
HasError := FConfigError OR (FResult = E_Result.Error);
END_GET
END_PROPERTY

{region 'Documentation'}
(*!
<summary>Reports a detected Reset timeout until Initialize or entry into a new Reset.</summary>
<description>
The owner leaves a timed-out Reset through Completing to Completed with Error, not through
Abort. Capacity waiting or scenario cleanup remains part of the configured deadline.
</description>
*)
{endregion}
{attribute 'monitoring' := 'call'}
PROPERTY PUBLIC HasResetTimeout : BOOL //! Reports a detected Reset timeout until Initialize or entry into a new Reset.
GET // PUBLIC
HasResetTimeout := FHasResetTimeout;
END_GET
END_PROPERTY

{region 'Documentation'}
(*!
<summary>Reports a detected execution timeout until Initialize or entry into a new Reset.</summary>
<description>
The owner supervises its own execution deadline; the parent does not duplicate this check.
Invalid timer measurements report Framework errors without setting this timeout flag.
</description>
*)
{endregion}
{attribute 'monitoring' := 'call'}
PROPERTY PUBLIC HasTimeout : BOOL //! Reports a detected execution timeout until Initialize or entry into a new Reset.
GET // PUBLIC
HasTimeout := FHasTimeout;
END_GET
END_PROPERTY

{region 'Documentation'}
(*!
<summary>Called by the PLC program after Event Buffer initialization and publisher
binding.</summary>
<description>
Name is validated before Configure. EventBuffer is retained and must match the selected
instance publisher. Rebuilds setup for PLC-start initialization; not an active-run recovery
operation. Success queues one initial Reset for the regular FB call; failure queues none.

Reinitialization requires configuration reactivation or PLC Cold Reset followed by the
application's first-cycle initialization chain. Normal PLC Stop/Start and UnitTest Reset do not
rebuild configuration. Do not call Initialize as recovery during an active run.

The selected publisher must already be usable for configuration diagnostics. Failure leaves
IsInitialized FALSE; retained diagnostic identity is not proof of valid setup.
</description>
*)
{endregion}
METHOD PUBLIC FINAL Initialize : BOOL //! TRUE after successful identity and setup validation; FALSE leaves the object uninitialized.
VAR_INPUT
    Name : STRING(2 * GVL_Constants.NameLength + 1); //! Nonempty root name without dots; validated before Configure and limited to NameLength.
    // SA0027: Parameter denotes the supplied service, not the EventBuffer FB type.
    {attribute 'analysis' := '-27'}
    EventBuffer : I_EventBuffer; //! Initialized buffer service retained for the Run Control lifetime; must match its selected event publisher.
END_VAR
VAR
    DefaultConfig : ST_RunConfig;
    EmptyStatus : ST_RunControlStatus;
    EmptyCollectionConfiguration : ST_TestSuiteCollectionConfig;
    // SA0167: Setup-only builder; no state or binding survives this initialization call.
    {attribute 'analysis' := '-167'}
    Builder : RunControlConfigurationBuilder;
    BufferStatus : ST_FifoStatus;
END_VAR
Initialize := FALSE;
FInitialized := FALSE;
FHasTimeout := FALSE;
FHasResetTimeout := FALSE;
FHasAbortTimeout := FALSE;
FCheckingInitialization := FALSE;
FConfigError := TRUE;
FEventBuffer := 0;
FCollectionConfiguration := EmptyCollectionConfiguration;
FConfig := DefaultConfig;
// SA0175: ASCII name contract; byte-based access is intentional and bounded.
{analysis -175}
FName := LEFT(Name, UINT_TO_INT(GVL_Constants.NameLength));
{analysis +175}
FResourceName := '';
FState := E_State.Uninitialized;
FResult := E_Result.NotEvaluated;
FStatus := EmptyStatus;
FExecutionTimer.Reset();
FStateTimer.Start();
FAggregator.Reset();
FTestSuiteCountInactive := 0;
FTestSuiteCountIdle := 0;
FTestSuiteCountRunning := 0;
FTestSuiteCountCompleted := 0;
FTestSuiteCountError := 0;
FCollectionValid := FALSE;
FChildrenError := FALSE;
FChildrenAborted := FALSE;
FChildrenCompleted := FALSE;
FChildrenAbortFinished := FALSE;
FFinalizationPublished := FALSE;
FMethodRequests.Start := FALSE;
FMethodRequests.Abort := FALSE;
FMethodRequests.Reset := FALSE;
UpdateStatus();

IF NOT IsNameValid(Name := Name, Depth := 1) THEN
    PublishInitializationError(Message := CONCAT('Invalid Run Control name: ', Name));
    RETURN;
END_IF;
IF EventBuffer = 0 THEN
    PublishInitializationError(Message := 'Missing Event Buffer interface.');
    RETURN;
END_IF;
IF NOT EventPublisher.IsValid THEN
    PublishInitializationError(Message := 'Event publisher is not ready for initialization.');
    RETURN;
END_IF;
BufferStatus := EventBuffer.FifoStatus;
IF BufferStatus.ConfigError OR BufferStatus.IndexError THEN
    PublishInitializationError(Message := 'Event Buffer configuration or indices are invalid.');
    RETURN;
END_IF;
FEventBuffer := EventBuffer;

Configure(Builder := Builder);
FCollectionConfiguration := Builder.Finalize();
IF NOT FCollectionConfiguration.IsValid THEN
    PublishInitializationError(Message := 'Invalid Test Suite collection configuration.');
    RETURN;
END_IF;

IF FOrchestrator = 0 THEN
    FOrchestrator := FDefaultOrchestrator;
END_IF;

FCheckingInitialization := TRUE;
IF NOT FOrchestrator.Initialize(Collection := THIS^,
    Name := FName,
    ResourceName := FResourceName) THEN
    FCheckingInitialization := FALSE;
    PublishInitializationError(Message := 'Orchestrator initialization failed.');
    UpdateStatus();
    RETURN;
END_IF;

FConfigError := NOT CheckInitialization();
FCheckingInitialization := FALSE;
IF FConfigError THEN
    UpdateStatus();
    RETURN;
END_IF;

FInitialized := TRUE;
RequestReset();
UpdateStatus();
Initialize := TRUE;
END_METHOD

{region 'Documentation'}
(*!
<summary>Reports completed explicit abort, including the legacy Aborted state.</summary>
*)
{endregion}
{attribute 'monitoring' := 'call'}
PROPERTY PUBLIC IsAborted : BOOL //! Reports completed explicit abort, including the legacy Aborted state.
GET // PUBLIC
IsAborted := ((FState = E_State.Completed) AND (FResult = E_Result.Abort)) OR (FState = E_State.Aborted);
END_GET
END_PROPERTY

{region 'Documentation'}
(*!
<summary>Reports explicit or error-driven abort processing.</summary>
*)
{endregion}
{attribute 'monitoring' := 'call'}
PROPERTY PUBLIC IsAborting : BOOL //! Reports explicit or error-driven abort processing.
GET // PUBLIC
IsAborting := (FState = E_State.Aborting) OR (FState = E_State.AbortingFromError);
END_GET
END_PROPERTY

{region 'Documentation'}
(*!
<summary>Reports terminal completion independently of the result.</summary>
*)
{endregion}
{attribute 'monitoring' := 'call'}
PROPERTY PUBLIC IsComplete : BOOL //! Reports terminal completion independently of the result.
GET // PUBLIC
IsComplete := FState = E_State.Completed;
END_GET
END_PROPERTY

{region 'Documentation'}
(*!
<summary>Reports completion-delay clock validity without modifying the timer; controlled test adapters may override this observation.</summary>
*)
{endregion}
{attribute 'monitoring' := 'call'}
PROPERTY PROTECTED IsCompletionTimeValid : BOOL //! Reports completion-delay clock validity without modifying the timer; controlled test adapters may override this observation.
GET
IsCompletionTimeValid := FStateTimer.IsValid;
END_GET
END_PROPERTY

{region 'Documentation'}
(*!
<summary>Reports Idle state independently of readiness.</summary>
*)
{endregion}
{attribute 'monitoring' := 'call'}
PROPERTY PUBLIC IsIdle : BOOL //! Reports Idle state independently of readiness.
GET // PUBLIC
IsIdle := FState = E_State.Idle;
END_GET
END_PROPERTY

{region 'Documentation'}
(*!
<summary>TRUE after successful configuration and child initialization checks.</summary>
*)
{endregion}
{attribute 'monitoring' := 'call'}
PROPERTY PUBLIC IsInitialized : BOOL //! TRUE after successful configuration and child initialization checks.
GET // PUBLIC
IsInitialized := FInitialized;
END_GET
END_PROPERTY

{region 'Documentation'}
(*!
<summary>Reports whether this owner can accept Start in Idle.</summary>
<description>
Requires successful initialization, valid configuration and collection, no owner Error, and
Orchestrator readiness with a neutral NotEvaluated helper result. The Orchestrator supplies the
child-readiness summary; IsInitialized or IsIdle alone is insufficient.
</description>
*)
{endregion}
{attribute 'monitoring' := 'call'}
PROPERTY PUBLIC IsReady : BOOL //! Reports whether this owner can accept Start in Idle.
GET // PUBLIC
IsReady := FALSE;
IF NOT FInitialized OR FConfigError OR (FResult = E_Result.Error) OR (FState <> E_State.Idle)
    OR NOT FCollectionValid THEN
    RETURN;
END_IF;
IsReady := FOrchestrator.IsReady
    AND (FOrchestrator.Result = E_Result.NotEvaluated);
END_GET
END_PROPERTY

{region 'Documentation'}
(*!
<summary>Reports active Reset processing.</summary>
*)
{endregion}
{attribute 'monitoring' := 'call'}
PROPERTY PUBLIC IsResetting : BOOL //! Reports active Reset processing.
GET // PUBLIC
IsResetting := FState = E_State.Reset;
END_GET
END_PROPERTY

{region 'Documentation'}
(*!
<summary>Reports the active lifecycle, including finalization and abort processing.</summary>
*)
{endregion}
{attribute 'monitoring' := 'call'}
PROPERTY PUBLIC IsRunControlActive : BOOL //! Reports the active lifecycle, including finalization and abort processing.
GET // PUBLIC
IsRunControlActive := (FState = E_State.Starting) OR (FState = E_State.Running)
    OR (FState = E_State.Completing) OR IsAborting;
END_GET
END_PROPERTY

{region 'Documentation'}
(*!
<summary>Checks a Run Control transition without changing state or producing diagnostics.</summary>
*)
{endregion}
METHOD PRIVATE IsStateTransitionAllowed : BOOL //! TRUE when NewState is allowed by the current initialization, lifecycle, readiness and completion conditions.
VAR_INPUT
    NewState : E_State; //! Requested lifecycle destination to check without changing state or emitting a diagnostic.
END_VAR
IF NewState = E_State.Uninitialized THEN
    IsStateTransitionAllowed := TRUE;
    RETURN;
END_IF;
IF NOT FInitialized THEN
    IsStateTransitionAllowed := FALSE;
    RETURN;
END_IF;

CASE NewState OF
    E_State.Reset:
        IsStateTransitionAllowed := TRUE;
    E_State.Idle:
        IsStateTransitionAllowed := (FState = E_State.Reset) AND NOT FConfigError
            AND (FResult <> E_Result.Error) AND FCollectionValid
            AND FOrchestrator.IsResetFinished
            AND (FOrchestrator.Result = E_Result.NotEvaluated);
    E_State.Starting:
        IsStateTransitionAllowed := IsReady;
    E_State.Running:
        IsStateTransitionAllowed := (FState = E_State.Starting) AND (FResult <> E_Result.Error);
    E_State.Completing:
        CASE FState OF
            E_State.Uninitialized, E_State.Starting, E_State.Completed:
                IsStateTransitionAllowed := FALSE;
            E_State.Reset, E_State.Idle:
                IsStateTransitionAllowed := FResult = E_Result.Error;
            E_State.Running:
                IsStateTransitionAllowed := FChildrenCompleted AND (FResult <> E_Result.Error)
                    AND FOrchestrator.IsExecutionFinished;
            E_State.Aborting, E_State.AbortingFromError:
                IsStateTransitionAllowed := TRUE;
        ELSE
            IsStateTransitionAllowed := FResult = E_Result.Error;
        END_CASE;
    E_State.Completed:
        IsStateTransitionAllowed := (FState = E_State.Completing) AND FFinalizationPublished
            AND (NOT IsCompletionTimeValid
                OR (FStateTimer.ElapsedLTime >= TIME_TO_LTIME(FConfig.CompletionDelay)));
    E_State.Aborting:
        IsStateTransitionAllowed := ((FState = E_State.Starting) OR (FState = E_State.Running))
            AND (FResult <> E_Result.Error);
    E_State.AbortingFromError:
        IsStateTransitionAllowed := ((FState = E_State.Starting) OR (FState = E_State.Running)
            OR (FState = E_State.Aborting)) AND (FResult = E_Result.Error);
ELSE
    IsStateTransitionAllowed := FALSE;
END_CASE;
END_METHOD

{region 'Documentation'}
(*!
<summary>Maps owner state and the current helper task; Reset finalization never selects Abort.</summary>
*)
{endregion}
METHOD PRIVATE MapOrchestratorTask : E_OrchestratorTask //! Helper task selected for State; Completing retains Execution/Abort, otherwise returns Idle.
VAR_INPUT
    State : E_State; //! Current owner lifecycle state after sequencing.
    CurrentTask : E_OrchestratorTask; //! Previously assigned helper task, retained during Completing only for Execution or Abort.
END_VAR
CASE State OF
    E_State.Reset:
        MapOrchestratorTask := E_OrchestratorTask.Reset;
    E_State.Starting, E_State.Running:
        MapOrchestratorTask := E_OrchestratorTask.Execution;
    E_State.Aborting, E_State.AbortingFromError:
        MapOrchestratorTask := E_OrchestratorTask.Abort;
    E_State.Completing:
        IF (CurrentTask = E_OrchestratorTask.Execution) OR (CurrentTask = E_OrchestratorTask.Abort) THEN
            MapOrchestratorTask := CurrentTask;
        ELSE
            MapOrchestratorTask := E_OrchestratorTask.Idle;
        END_IF;
ELSE
    MapOrchestratorTask := E_OrchestratorTask.Idle;
END_CASE;
END_METHOD

{region 'Documentation'}
(*!
<summary>Root identity retained for diagnostics, including rejected names.</summary>
*)
{endregion}
{attribute 'monitoring' := 'variable'}
PROPERTY PUBLIC Name : STRING(GVL_Constants.NameLength) //! Root identity retained for diagnostics, including rejected names.
GET // PUBLIC
Name := FName;
END_GET
END_PROPERTY

{region 'Documentation'}
(*!
<summary>Reads one child snapshot and accumulates lifecycle observations; invalid bindings invalidate the collection.</summary>
*)
{endregion}
METHOD PRIVATE ObserveTestSuite : BOOL //! TRUE after reading an initialized child snapshot; FALSE clears ChildStatus and invalidates collection observations.
VAR_INPUT
    Child : I_TestSuite; //! Borrowed Suite interface; zero or uninitialized children invalidate the collection observations.
END_VAR
VAR_OUTPUT
    ChildStatus : ST_TestSuiteStatus; //! One child snapshot by value; default empty status on invalid binding. TRUE is binding validity, not a successful test result.
END_VAR
VAR
    ChildValid : BOOL;
    EmptyStatus : ST_TestSuiteStatus;
END_VAR
ObserveTestSuite := FALSE;
ChildValid := FALSE;
IF Child <> 0 THEN
    ChildValid := Child.IsInitialized;
END_IF;
IF NOT ChildValid THEN
    ChildStatus := EmptyStatus;
    FCollectionValid := FALSE;
    FChildrenCompleted := FALSE;
    FChildrenAbortFinished := FALSE;
    FChildrenError := TRUE;
    RETURN;
END_IF;

ChildStatus := Child.Status;
CASE ChildStatus.Execution.Result OF
    E_Result.NotEvaluated, E_Result.Passed, E_Result.Failed, E_Result.Abort, E_Result.Error:
        FChildrenError := FChildrenError OR (ChildStatus.Execution.Result = E_Result.Error);
ELSE
    FChildrenError := TRUE;
END_CASE;
FChildrenError := FChildrenError OR ChildStatus.Execution.Error OR ChildStatus.Execution.ConfigError
    OR (ChildStatus.Execution.ExecutionStatus = E_ExecutionStatus.Error);
FChildrenAborted := FChildrenAborted OR (ChildStatus.Execution.Result = E_Result.Abort);
FChildrenCompleted := FChildrenCompleted AND ChildStatus.Execution.Completed;
FChildrenAbortFinished := FChildrenAbortFinished
    AND (ChildStatus.Execution.Ready OR ChildStatus.Execution.Completed);
ObserveTestSuite := TRUE;
END_METHOD

{region 'Documentation'}
(*!
<summary>Processes Buffer commands before lifecycle work; Reset follows every hierarchical release attempt.</summary>
<description>
Release return values do not gate the hard reset. Delete retains the external field's snapshot semantics.
</description>
*)
{endregion}
METHOD PRIVATE ProcessBufferCommands
VAR_IN_OUT
    Commands : ST_EventBufferCommand; //! Actual external Buffer command storage; Reset releases reservations then clears both commands; Delete uses captured watermark semantics.
END_VAR
VAR
    Index : LINT;
    Child : I_TestSuite;
END_VAR
IF FEventBuffer = 0 THEN
    RETURN;
END_IF;

IF Commands.Reset THEN
    FOR Index := DINT_TO_LINT(ChildArrayLowerBound) TO DINT_TO_LINT(ChildArrayLowerBound) + UINT_TO_LINT(ChildCount) - 1 DO
        Child := GetTestSuite(Index := LINT_TO_DINT(Index));
        IF Child <> 0 THEN
            Child.FreeReservedEvents();
        END_IF;
    END_FOR;

    FEventBuffer.Reset();
    Commands.Reset := FALSE;
    Commands.DeleteSequenceId := 0;
    RETURN;
END_IF;

FEventBuffer.ProcessDeleteRequest(SequenceId := Commands.DeleteSequenceId);
END_METHOD

{region 'Documentation'}
(*!
<summary>Consumes same-task requests, reports each received request and prioritizes Reset &gt; Abort &gt; Start.</summary>
<description>
Discards requests before initialization; never changes lifecycle state.
</description>
*)
{endregion}
METHOD PRIVATE ProcessRequests
VAR_IN_OUT
    InputRequests : ST_Command; //! Same-task request mailbox consumed and cleared by this call, including before initialization.
END_VAR
VAR_OUTPUT
    Requests : ST_Command; //! Qualified request snapshot with Reset over Abort over Start; all FALSE before initialization.
END_VAR
Requests.Reset := FALSE;
Requests.Abort := FALSE;
Requests.Start := FALSE;

IF NOT FInitialized THEN
    InputRequests.Reset := FALSE;
    InputRequests.Abort := FALSE;
    InputRequests.Start := FALSE;
    RETURN;
END_IF;

Requests.Reset := InputRequests.Reset;
Requests.Abort := InputRequests.Abort AND NOT InputRequests.Reset;
Requests.Start := InputRequests.Start AND NOT InputRequests.Abort AND NOT InputRequests.Reset;

IF InputRequests.Reset THEN
    PublishEvent(Event := CreateResetEvent(OwnerScope := E_OwnerScope.RunControl,
        Name := FName,
        ResourceName := FResourceName,
        State := FState));
END_IF;

IF InputRequests.Abort THEN
    PublishEvent(Event := CreateAbortEvent(OwnerScope := E_OwnerScope.RunControl,
        Name := FName,
        ResourceName := FResourceName,
        State := FState));
END_IF;

IF InputRequests.Start THEN
    PublishEvent(Event := CreateStartEvent(OwnerScope := E_OwnerScope.RunControl,
        Name := FName,
        ResourceName := FResourceName,
        State := FState));
END_IF;

InputRequests.Reset := FALSE;
InputRequests.Abort := FALSE;
InputRequests.Start := FALSE;
END_METHOD

{region 'Documentation'}
(*!
<summary>Calls every owned Suite exactly once per initialized cycle, including Completed.</summary>
<description>
Do not gate child calls by parent state; child requests and lifecycle control their
work.
</description>
*)
{endregion}
METHOD PROTECTED ABSTRACT ProcessTestSuites
(* Example: call every owned Suite, including children not currently selected.
FTestSuiteA();
FTestSuiteB();
*)
END_METHOD

{region 'Documentation'}
(*!
<summary>Publishes through the selected instance publisher without owning buffer loss accounting.</summary>
*)
{endregion}
METHOD PRIVATE PublishEvent
VAR_INPUT
    Event : ST_Event; //! Payload value forwarded once to the selected publisher; the publisher assigns identity/time and accounts for loss.
END_VAR
EventPublisher.PublishEvent(Event := Event);
END_METHOD

{region 'Documentation'}
(*!
<summary>Emits a setup diagnostic through the required usable selected publisher; leaves lifecycle and result unchanged.</summary>
*)
{endregion}
METHOD PRIVATE PublishInitializationError
VAR_INPUT
    Message : STRING(GVL_Constants.MessageLength); //! Setup diagnostic text sent through the required usable selected publisher; lifecycle and result are unchanged.
END_VAR
EventPublisher.PublishEvent(Event := CreateFrameworkEvent(Name := FName,
    ResourceName := FResourceName,
    State := E_State.Uninitialized,
    Severity := E_EventSeverity.Error,
    Message := Message));
END_METHOD

{region 'Documentation'}
(*!
<summary>Records an Abort request for the next regular FB call.</summary>
<description>
Repeated positive calls coalesce in the same-task request storage. Processing consumes the
requests with priority Reset, Abort, Start; calls before successful initialization are discarded
when processed.

Abort requests controlled termination of execution, not Reset cancellation. The owner
lifecycle determines whether the request applies.
</description>
*)
{endregion}
METHOD PUBLIC RequestAbort
FMethodRequests.Abort := TRUE;
END_METHOD

{region 'Documentation'}
(*!
<summary>Records a Reset request for the next regular FB call.</summary>
<description>
Repeated positive calls coalesce in the same-task request storage. Processing consumes the
requests with priority Reset, Abort, Start; calls before successful initialization are discarded
when processed.

Lifecycle Reset preserves configuration and publisher binding. It is not reinitialization or
Event Buffer Reset.
</description>
*)
{endregion}
METHOD PUBLIC RequestReset
FMethodRequests.Reset := TRUE;
END_METHOD

{region 'Documentation'}
(*!
<summary>Records a Start request for the next regular FB call.</summary>
<description>
Repeated positive calls coalesce in the same-task request storage. Processing consumes the
requests with priority Reset, Abort, Start; calls before successful initialization are discarded
when processed.

Start is accepted by the lifecycle only in ready Idle. Recording the request does not start
execution synchronously.
</description>
*)
{endregion}
METHOD PUBLIC RequestStart
FMethodRequests.Start := TRUE;
END_METHOD

{region 'Documentation'}
(*!
<summary>Current owner result; final publication holds it until Reset or explicit
initialization.</summary>
*)
{endregion}
{attribute 'monitoring' := 'call'}
PROPERTY PUBLIC Result : E_Result //! Current owner result; final publication holds it until Reset or explicit initialization.
GET // PUBLIC
Result := FResult;
END_GET
END_PROPERTY

{region 'Documentation'}
(*!
<summary>Owns Run Control transition decisions; child dispatch belongs to the shared Orchestrator.</summary>
*)
{endregion}
METHOD PRIVATE Sequencer
VAR_INPUT
    Requests : ST_Command; //! Consumed lifecycle request snapshot; transition applicability is checked against the current owner state.
END_VAR
IF NOT FInitialized THEN
    IF FState <> E_State.Uninitialized THEN
        ChangeState(NewState := E_State.Uninitialized);
    END_IF;
    RETURN;
END_IF;
IF Requests.Reset THEN
    ChangeState(NewState := E_State.Reset);
END_IF;

CASE FState OF
    E_State.Uninitialized:
        RETURN;

    E_State.Reset:
        IF NOT FStateTimer.IsValid THEN
            Error(Message := 'Task clock error during Run Control reset.');
            ChangeState(NewState := E_State.Completing);
            RETURN;
        END_IF;
        IF FStateTimer.ElapsedLTime >= TIME_TO_LTIME(FConfig.ResetTimeout) THEN
            FHasResetTimeout := TRUE;
            PublishEvent(Event := CreateFrameworkEvent(Name := FName,
                ResourceName := FResourceName,
                State := FState,
                Severity := E_EventSeverity.Error,
                Message := 'Run Control reset timeout reached.'));
            FResult := E_Result.Error;
            ChangeState(NewState := E_State.Completing);
            RETURN;
        END_IF;
        IF NOT FOrchestrator.IsResetActive THEN
            RETURN;
        END_IF;
        IF NOT FCollectionValid THEN
            Error(Message := 'Registered Test Suite collection is no longer valid.');
            ChangeState(NewState := E_State.Completing);
            RETURN;
        END_IF;
        IF FOrchestrator.Result = E_Result.Error THEN
            Error(Message := 'Orchestrator failed during Run Control reset.');
        END_IF;
        IF (FResult = E_Result.Error) AND FOrchestrator.IsResetFinished THEN
            ChangeState(NewState := E_State.Completing);
            RETURN;
        END_IF;
        IF FOrchestrator.IsResetFinished THEN
            ChangeState(NewState := E_State.Idle);
        END_IF;
        RETURN;

    E_State.Idle:
        IF FResult = E_Result.Error THEN
            ChangeState(NewState := E_State.Completing);
            RETURN;
        END_IF;
        IF Requests.Start AND IsReady THEN
            ChangeState(NewState := E_State.Starting);
        END_IF;
        RETURN;

    E_State.Starting, E_State.Running:
        IF NOT FCollectionValid THEN
            Error(Message := 'Registered Test Suite collection is no longer valid.');
            ChangeState(NewState := E_State.AbortingFromError);
            RETURN;
        END_IF;
        IF FResult <> E_Result.Error THEN
            IF FChildrenError THEN
                Error(Message := 'A registered Test Suite reported an error.');
            ELSIF FChildrenAborted AND (FResult <> E_Result.Abort) THEN
                Error(Message := 'Unexpected Test Suite abort.');
            END_IF;
        END_IF;
        IF FResult = E_Result.Error THEN
            ChangeState(NewState := E_State.AbortingFromError);
            RETURN;
        END_IF;
        IF FOrchestrator.Result = E_Result.Error THEN
            Error(Message := 'Orchestrator reported an execution error.');
            ChangeState(NewState := E_State.AbortingFromError);
            RETURN;
        END_IF;
        IF NOT FExecutionTimer.IsValid THEN
            Error(Message := 'Task clock error during Run Control execution.');
            ChangeState(NewState := E_State.AbortingFromError);
            RETURN;
        END_IF;
        IF FExecutionTimer.ElapsedLTime >= TIME_TO_LTIME(FConfig.Timeout) THEN
            FHasTimeout := TRUE;
            Error(Message := 'Run Control timeout reached.');
            ChangeState(NewState := E_State.AbortingFromError);
            RETURN;
        END_IF;
        IF Requests.Abort THEN
            ChangeState(NewState := E_State.Aborting);
            RETURN;
        END_IF;
        IF FState = E_State.Starting THEN
            ChangeState(NewState := E_State.Running);
            RETURN;
        END_IF;
        IF FChildrenCompleted AND FOrchestrator.IsExecutionFinished THEN
            ChangeState(NewState := E_State.Completing);
        END_IF;
        RETURN;

    E_State.Completing:
        IF FFinalizationPublished AND NOT IsCompletionTimeValid THEN
            PublishEvent(Event := CreateFrameworkEvent(Name := FName,
                ResourceName := FResourceName,
                State := FState,
                Severity := E_EventSeverity.Error,
                Message := 'Task clock error during Run Control completion delay.'));
            ChangeState(NewState := E_State.Completed);
            RETURN;
        END_IF;
        IF FFinalizationPublished AND (FStateTimer.ElapsedLTime >= TIME_TO_LTIME(FConfig.CompletionDelay)) THEN
            ChangeState(NewState := E_State.Completed);
        END_IF;
        RETURN;

    E_State.Completed:
        RETURN;

    E_State.Aborting, E_State.AbortingFromError:
        IF (FState = E_State.Aborting) AND NOT FCollectionValid THEN
            Error(Message := 'Registered Test Suite collection is no longer valid.');
            ChangeState(NewState := E_State.AbortingFromError);
            RETURN;
        END_IF;
        IF FResult <> E_Result.Error THEN
            IF FChildrenError THEN
                Error(Message := 'A registered Test Suite reported an error.');
            ELSIF FChildrenAborted AND (FResult <> E_Result.Abort) AND (FState <> E_State.Aborting) THEN
                Error(Message := 'Unexpected Test Suite abort.');
            END_IF;
        END_IF;
        IF NOT FStateTimer.IsValid THEN
            PublishEvent(Event := CreateFrameworkEvent(Name := FName,
                ResourceName := FResourceName,
                State := FState,
                Severity := E_EventSeverity.Error,
                Message := 'Task clock error during Run Control abort.'));
            FResult := E_Result.Error;
            ChangeState(NewState := E_State.Completing);
            RETURN;
        END_IF;
        IF FStateTimer.ElapsedLTime >= TIME_TO_LTIME(FConfig.AbortTimeout) THEN
            FHasAbortTimeout := TRUE;
            PublishEvent(Event := CreateFrameworkEvent(Name := FName,
                ResourceName := FResourceName,
                State := FState,
                Severity := E_EventSeverity.Error,
                Message := 'Run Control abort timeout reached.'));
            FResult := E_Result.Error;
            ChangeState(NewState := E_State.Completing);
            RETURN;
        END_IF;
        IF (FState = E_State.Aborting) AND (FResult = E_Result.Error) THEN
            ChangeState(NewState := E_State.AbortingFromError);
            RETURN;
        END_IF;
        IF (FState = E_State.Aborting)
            AND (FOrchestrator.Result = E_Result.Error) THEN
            Error(Message := 'Orchestrator failed during Run Control abort.');
            ChangeState(NewState := E_State.AbortingFromError);
            RETURN;
        END_IF;
        IF FChildrenAbortFinished AND FOrchestrator.IsAbortFinished THEN
            ChangeState(NewState := E_State.Completing);
        END_IF;
        RETURN;
ELSE
    Error(Message := 'Unhandled Run Control lifecycle state.');
    ChangeState(NewState := E_State.Completing);
END_CASE;
END_METHOD

{region 'Documentation'}
(*!
<summary>Current Run Control lifecycle state.</summary>
*)
{endregion}
{attribute 'monitoring' := 'call'}
PROPERTY PUBLIC State : E_State //! Current Run Control lifecycle state.
GET // PUBLIC
State := FState;
END_GET
END_PROPERTY

{region 'Documentation'}
(*!
<summary>Returns the latest cyclic owner-status snapshot.</summary>
<description>
Status is refreshed on every FB call, including Uninitialized and Completed. Runtime uses
TIME; child counters may continue changing after final event publication. Reading this property
performs no child processing and does not republish final events.
</description>
*)
{endregion}
{attribute 'monitoring' := 'variable'}
PROPERTY PUBLIC Status : ST_RunControlStatus //! Returns the latest cyclic owner-status snapshot.
GET // PUBLIC
Status := FStatus;
END_GET
END_PROPERTY

{region 'Documentation'}
(*!
<summary>Applies owner result semantics to the current child aggregate without changing lifecycle state.</summary>
*)
{endregion}
METHOD PRIVATE UpdateResult
VAR
    OrchestratorResult : E_Result;
END_VAR
IF FState = E_State.Uninitialized THEN
    FResult := E_Result.NotEvaluated;
    RETURN;
END_IF;
IF (FState = E_State.Reset) OR (FState = E_State.Completed) OR FFinalizationPublished
    OR (FResult = E_Result.Error) THEN
    RETURN;
END_IF;

IF NOT FCollectionValid THEN
    Error(Message := 'Registered Test Suite collection is no longer valid.');
    RETURN;
END_IF;
IF FChildrenError OR (FAggregator.Result = E_Result.Error) THEN
    Error(Message := 'A registered Test Suite reported an error.');
    RETURN;
END_IF;
OrchestratorResult := FOrchestrator.Result;
IF OrchestratorResult = E_Result.Error THEN
    Error(Message := 'Orchestrator reported an error.');
    RETURN;
END_IF;
IF (FAggregator.Result = E_Result.Abort)
    AND (FResult <> E_Result.Abort) AND (FState <> E_State.Aborting) THEN
    Error(Message := 'Unexpected Test Suite abort.');
    RETURN;
END_IF;

CASE FState OF
    E_State.Idle, E_State.Starting, E_State.Running:
        FResult := E_Result.NotEvaluated;
    E_State.Aborting:
        FResult := E_Result.Abort;
    E_State.AbortingFromError:
        FResult := E_Result.Error;
    E_State.Completing:
        IF FResult = E_Result.Abort THEN
            RETURN;
        END_IF;
        IF (FResult = E_Result.Failed) OR (FAggregator.Result = E_Result.Failed) THEN
            FResult := E_Result.Failed;
            RETURN;
        END_IF;
        FResult := E_Result.Passed;
ELSE
    Error(Message := 'Unhandled Run Control lifecycle state.');
END_CASE;
END_METHOD

{region 'Documentation'}
(*!
<summary>Projects lifecycle, runtime and internally collected counters on every FB call, including Completed.</summary>
*)
{endregion}
METHOD PRIVATE UpdateStatus
VAR
    Execution : ST_ExecutionStatus;
END_VAR
Execution.State := FState;
Execution.Result := FResult;
Execution.ConfigError := FConfigError;
CASE FState OF
    E_State.Uninitialized:
        Execution.ExecutionStatus := E_ExecutionStatus.NotReady;
        Execution.Uninitialized := TRUE;
    E_State.Reset:
        Execution.ExecutionStatus := E_ExecutionStatus.Reset;
    E_State.Idle:
        Execution.ExecutionStatus := E_ExecutionStatus.Idle;
        Execution.Ready := IsReady;
    E_State.Starting:
        Execution.ExecutionStatus := E_ExecutionStatus.Starting;
    E_State.Running:
        Execution.ExecutionStatus := E_ExecutionStatus.Running;
        Execution.Running := TRUE;
    E_State.Completing:
        Execution.ExecutionStatus := E_ExecutionStatus.Completing;
    E_State.Completed:
        Execution.ExecutionStatus := E_ExecutionStatus.Completed;
        Execution.Completed := TRUE;
        Execution.Aborted := FResult = E_Result.Abort;
    E_State.Aborting, E_State.AbortingFromError:
        Execution.ExecutionStatus := E_ExecutionStatus.Aborting;
ELSE
    Execution.ExecutionStatus := E_ExecutionStatus.Error;
END_CASE;
Execution.Error := HasError;
FStatus.Execution := Execution;
FStatus.Runtime := FExecutionTimer.ElapsedTime;
FStatus.SuiteCountTotal := ChildCount;
FStatus.SuiteCountInactive := FTestSuiteCountInactive;
FStatus.SuiteCountIdle := FTestSuiteCountIdle;
FStatus.SuiteCountRunning := FTestSuiteCountRunning;
FStatus.SuiteCountCompleted := FTestSuiteCountCompleted;
FStatus.SuiteCountError := FTestSuiteCountError;
FStatus.SuiteCountPassed := FAggregator.PassedCount;
FStatus.SuiteCountFailed := FAggregator.FailedCount;
END_METHOD

END_FUNCTION_BLOCK

// ---- Framework/Common/POU/Orchestrator.TcPOU
{region 'Documentation'}
(*!
<summary>Owner-driven child slot scheduler; call before concrete children, once per task cycle.</summary>
<description>
The owner supplies a validated nonempty collection with a contiguous occupied prefix and ordered execution slots. Collection bounds, children and slots remain fixed until full reinitialization; Initialize caches occupied indices rather than validating array capacity again. Keep the collection, children and selected publisher alive. Use either the concrete FB call or Execute once per cycle, before the owner calls every concrete child; this helper never calls child FB bodies, aggregates child results or supervises owner timeouts.

Execution starts at slot one. At most one fitting child Start is requested per call; capacity-waiting candidates may be skipped within a shared slot. A later slot waits for all children in the current slot to complete. Reset dispatch is independent of execution slots and admits at most one new Reset per call, allowing admitted resets to overlap. Reservations are acquired through the child before each request and released through its owner operation at the applicable stable boundary.

Repeating the same task preserves progress. Task completion never changes the assigned task. Technical Error blocks new execution Starts but does not cancel remaining Reset attempts; it is held through Idle and Abort until Initialize or entry into a new Reset task. Completion and success are separate: Reset or Abort can finish with Error. The owner decides the lifecycle reaction and must continue concrete child calls, including after owner completion. Processing scans the registered children and may invoke hierarchical releases; cost depends on the configured collection and subtree.
</description>
*)
{endregion}
FUNCTION_BLOCK Orchestrator IMPLEMENTS I_Orchestrator
VAR_INPUT
    Task : E_OrchestratorTask := E_OrchestratorTask.Idle; //! Owner-selected task, supplied on every cyclic call.
END_VAR
VAR
    /// Instance binding; derived test adapters may assign it before first use.
    FEventPublisher : I_EventPublisher;
    FCollection : I_OrchestratableCollection;
    FInitialized : BOOL;
    FFirstOccupiedIndex : DINT;
    FName : STRING(GVL_Constants.NameLength);
    FResourceName : STRING(GVL_Constants.ResourceNameLength);
    FResult : E_Result := E_Result.NotEvaluated;
    FPreviousTask : E_OrchestratorTask := E_OrchestratorTask.Idle;
    FResetFinished : BOOL;
    FAbortFinished : BOOL;
    FExecutionFinished : BOOL;
    FChildrenReady : BOOL;
    FLastOccupiedIndex : DINT;
    FNextResetOffset : UDINT;
    FCurrentSlot : UINT;
    FSlotFirstIndex : DINT;
    FSlotLastIndex : DINT;
    FHasPendingStart : BOOL;
    FPendingStartIndex : DINT;
END_VAR

IF NOT FInitialized THEN
    RETURN;
END_IF;

IF Task <> FPreviousTask THEN
    InitializeTask();
    FPreviousTask := Task;
END_IF;

CASE Task OF
    E_OrchestratorTask.Idle:
        ProcessIdle();
    E_OrchestratorTask.Reset:
        ProcessReset();
    E_OrchestratorTask.Execution:
        ProcessExecution();
    E_OrchestratorTask.Abort:
        ProcessAbort();
ELSE
    Error(Message := 'Unknown Orchestrator task.');
END_CASE;

{region 'Documentation'}
(*!
<summary>Requests controlled abort only from children not already stopped or aborting.</summary>
*)
{endregion}
METHOD PRIVATE AbortChildren
VAR
    Index : LINT;
    Child : I_Orchestratable;
END_VAR
FOR Index := DINT_TO_LINT(FFirstOccupiedIndex) TO DINT_TO_LINT(FLastOccupiedIndex) DO
    Child := ReadChild(Index := LINT_TO_DINT(Index));
    IF Child = 0 THEN
        CONTINUE;
    END_IF;
    IF (Child.State = E_State.Completed)
        OR ((Child.State = E_State.Idle) AND Child.IsReady)
        OR (Child.State = E_State.Aborting)
        OR (Child.State = E_State.AbortingFromError) THEN
        CONTINUE;
    END_IF;
    Child.RequestAbort();
END_FOR;
END_METHOD

{region 'Documentation'}
(*!
<summary>Selected unfinished Execution slot; zero when no Execution slot is active.</summary>
*)
{endregion}
{attribute 'monitoring' := 'call'}
PROPERTY PUBLIC ActiveSlot : UINT //! Selected unfinished Execution slot; zero when no Execution slot is active.
GET // PUBLIC
ActiveSlot := 0;
IF IsExecutionActive AND NOT IsExecutionFinished THEN
    ActiveSlot := FCurrentSlot;
END_IF;
END_GET
END_PROPERTY

{region 'Documentation'}
(*!
<summary>Checks child bindings, task-specific failures and current-slot invariants; latches diagnostics only.</summary>
*)
{endregion}
METHOD PRIVATE CheckChildErrors
VAR
    Index : LINT;
    Child : I_Orchestratable;
END_VAR
FOR Index := DINT_TO_LINT(FFirstOccupiedIndex) TO DINT_TO_LINT(FLastOccupiedIndex) DO
    Child := ReadChild(Index := LINT_TO_DINT(Index));
    IF Child = 0 THEN
        CONTINUE;
    END_IF;

    CASE Task OF
        E_OrchestratorTask.Reset:
            IF Index >= DINT_TO_LINT(FFirstOccupiedIndex) + UDINT_TO_LINT(FNextResetOffset) THEN
                CONTINUE;
            END_IF;
            IF Child.HasError
                OR ((Child.State = E_State.Completed) AND Child.IsComplete) THEN
                Error(Message := CONCAT('Child reset failed: ', Child.Name));
            END_IF;

        E_OrchestratorTask.Execution, E_OrchestratorTask.Abort:
            IF Child.HasError THEN
                Error(Message := CONCAT('Child reported an error: ', Child.Name));
            END_IF;
            IF (Task = E_OrchestratorTask.Execution) AND (Child.Result = E_Result.Abort) THEN
                Error(Message := CONCAT('Unexpected child Abort: ', Child.Name));
            END_IF;
    ELSE
        CONTINUE;
    END_CASE;

    IF (Task <> E_OrchestratorTask.Execution) OR (FCurrentSlot = 0)
        OR (Index < DINT_TO_LINT(FSlotFirstIndex)) OR (Index > DINT_TO_LINT(FSlotLastIndex)) THEN
        CONTINUE;
    END_IF;
    IF Child.ExecutionSlot <> FCurrentSlot THEN
        Error(Message := 'Child slot changed during execution.');
    END_IF;
    CASE Child.State OF
        E_State.Completed:
            IF NOT Child.IsComplete THEN
                Error(Message := CONCAT('Inconsistent child completion: ', Child.Name));
            END_IF;
        E_State.Idle:
            IF NOT Child.IsReady THEN
                Error(Message := CONCAT('Child is not ready for Start: ', Child.Name));
            END_IF;
        E_State.Starting..E_State.Completing:
            IF Child.ReservedEntryCount = 0 THEN
                Error(Message := CONCAT('Active child has no event reservation: ', Child.Name));
            END_IF;
    ELSE
        Error(Message := CONCAT('Unexpected child execution state: ', Child.Name));
    END_CASE;
END_FOR;
END_METHOD

{region 'Documentation'}
(*!
<summary>Checks the Child response to the previous Start; a missing reaction releases its reservation.</summary>
*)
{endregion}
METHOD PRIVATE CheckChildStarted
VAR_INPUT
    ChildIndex : DINT; //! Original collection index of the child whose previously dispatched Start is awaiting confirmation.
END_VAR
VAR_IN_OUT
    HasPendingStart : BOOL; //! TRUE while a previous Start awaits confirmation; cleared when that response is checked.
END_VAR
VAR
    Child : I_Orchestratable;
END_VAR
IF (Task = E_OrchestratorTask.Reset) OR NOT HasPendingStart THEN
    RETURN;
END_IF;
HasPendingStart := FALSE;
Child := ReadChild(Index := ChildIndex);
IF Child = 0 THEN
    RETURN;
END_IF;

IF Child.State = E_State.Idle THEN
    IF NOT Child.FreeReservedEvents() THEN
        Error(Message := CONCAT('Cannot release rejected Start reservation: ', Child.Name));
        RETURN;
    END_IF;
    Error(Message := CONCAT('Child did not react to Start: ', Child.Name));
    RETURN;
END_IF;
IF (Child.State = E_State.Uninitialized) OR (Child.State = E_State.Reset) THEN
    Error(Message := CONCAT('Unexpected state after child Start: ', Child.Name));
END_IF;
END_METHOD

{region 'Documentation'}
(*!
<summary>Last task supplied to the scheduler.</summary>
*)
{endregion}
{attribute 'monitoring' := 'call'}
PROPERTY PUBLIC CurrentTask : E_OrchestratorTask //! Last task supplied to the scheduler.
GET // PUBLIC
CurrentTask := Task;
END_GET
END_PROPERTY

{region 'Documentation'}
(*!
<summary>Latches the technical error and publishes its first diagnostic; never changes the supplied task.</summary>
*)
{endregion}
METHOD PRIVATE Error
VAR_INPUT
    Message : STRING(GVL_Constants.MessageLength); //! Technical diagnostic text published when this call first latches Error.
END_VAR
IF FResult = E_Result.Error THEN
    RETURN;
END_IF;
FResult := E_Result.Error;
PublishEvent(Event := CreateFrameworkEvent(Name := CONCAT(FName, '.Orchestrator'),
    ResourceName := FResourceName,
    State := E_State.Error,
    Severity := E_EventSeverity.Error,
    Message := Message));
END_METHOD

{region 'Documentation'}
(*!
<summary>Returns the retained instance service; binds the default only on first use.</summary>
*)
{endregion}
{attribute 'monitoring' := 'variable'}
PROPERTY PUBLIC EventPublisher : I_EventPublisher //! Returns the retained instance service; binds the default only on first use.
GET // PUBLIC
IF FEventPublisher = 0 THEN
    FEventPublisher := GVL_EventBuffer.Publisher;
END_IF;
EventPublisher := FEventPublisher;
END_GET
END_PROPERTY

{region 'Documentation'}
(*!
<summary>Executes the existing FB body once through the owner-facing interface.</summary>
*)
{endregion}
METHOD PUBLIC Execute
VAR_INPUT
    Task : E_OrchestratorTask; //! Owner-selected work for this call; a task change initializes its scheduling once.
END_VAR
THIS^(Task := Task);
END_METHOD

{region 'Documentation'}
(*!
<summary>Releases eligible child reservations before completion/admission; FALSE means at least one unresolved access or release.</summary>
*)
{endregion}
METHOD PRIVATE FreeCompletedReservations : BOOL //! TRUE when all eligible releases and required child accesses succeeded; FALSE permits partial release.
VAR
    Index : LINT;
    Child : I_Orchestratable;
    ReleaseReservation : BOOL;
END_VAR
FreeCompletedReservations := TRUE;
FOR Index := DINT_TO_LINT(FFirstOccupiedIndex) TO DINT_TO_LINT(FLastOccupiedIndex) DO
    Child := ReadChild(Index := LINT_TO_DINT(Index));
    IF Child = 0 THEN
        FreeCompletedReservations := FALSE;
        CONTINUE;
    END_IF;

    CASE Task OF
        E_OrchestratorTask.Reset:
            ReleaseReservation := (Child.State = E_State.Idle) AND Child.IsReady;
        E_OrchestratorTask.Execution:
            ReleaseReservation := (Child.State = E_State.Completed) AND Child.IsComplete;
        E_OrchestratorTask.Abort, E_OrchestratorTask.Idle:
            ReleaseReservation := ((Child.State = E_State.Idle) AND Child.IsReady)
                OR ((Child.State = E_State.Completed) AND Child.IsComplete);
    ELSE
        ReleaseReservation := FALSE;
    END_CASE;
    IF NOT ReleaseReservation THEN
        CONTINUE;
    END_IF;
    IF NOT Child.FreeReservedEvents() THEN
        Error(Message := CONCAT('Cannot release child reservation: ', Child.Name));
        FreeCompletedReservations := FALSE;
    END_IF;
END_FOR;
END_METHOD

{region 'Documentation'}
(*!
<summary>Binds the owner&#x27;s validated collection and caches its occupied bounds once. Clears scheduling state without calling children or changing their reservations.</summary>
<description>
This accepts a nonzero collection, nonempty Name and positive ChildCount, then caches the lower bound and occupied end. Capacity, naming and ordered slots are validated by the owner/builder. The owner also checks child initialization before enabling regular execution; this method does not repeat those checks. It drops the previous collection before validation, so a failed call leaves the helper uninitialized. Reinitialization is configuration setup, not active-run recovery.
</description>
*)
{endregion}
METHOD PUBLIC Initialize : BOOL //! TRUE when the child collection is accepted and scheduling is initialized.
VAR_INPUT
    Collection : I_OrchestratableCollection; //! Initialized, stable child collection retained by the scheduler; its owner and children must outlive use.
    Name : STRING(GVL_Constants.NameLength); //! Hierarchical owner name used to identify events; must satisfy the naming contract.
    ResourceName : STRING(GVL_Constants.ResourceNameLength) := ''; //! Optional resource context for diagnostics; empty by default.
END_VAR
VAR
    Count : UINT;
END_VAR
Initialize := FALSE;
FInitialized := FALSE;
FCollection := 0;
FFirstOccupiedIndex := 0;
FLastOccupiedIndex := 0;
FName := Name;
FResourceName := ResourceName;
FResult := E_Result.NotEvaluated;
Task := E_OrchestratorTask.Idle;
FPreviousTask := E_OrchestratorTask.Idle;
FResetFinished := FALSE;
FAbortFinished := FALSE;
FExecutionFinished := FALSE;
FChildrenReady := FALSE;
FNextResetOffset := 0;
FCurrentSlot := 0;
FSlotFirstIndex := 0;
FSlotLastIndex := 0;
FHasPendingStart := FALSE;
FPendingStartIndex := 0;

IF (Collection = 0) OR (Name = '') THEN
    RETURN;
END_IF;
Count := Collection.ChildCount;
IF Count = 0 THEN
    RETURN;
END_IF;

FFirstOccupiedIndex := Collection.ChildArrayLowerBound;
FLastOccupiedIndex := LINT_TO_DINT(DINT_TO_LINT(FFirstOccupiedIndex) + UINT_TO_LINT(Count) - 1);
FCollection := Collection;
FInitialized := TRUE;
Initialize := TRUE;
END_METHOD

{region 'Documentation'}
(*!
<summary>Initializes progress once when the supplied task changes; never selects another task.</summary>
*)
{endregion}
METHOD PRIVATE InitializeTask
CASE Task OF
    E_OrchestratorTask.Idle:
        FHasPendingStart := FALSE;

    E_OrchestratorTask.Reset:
        FCurrentSlot := 0;
        FNextResetOffset := 0;
        FHasPendingStart := FALSE;
        FResult := E_Result.NotEvaluated;
        FResetFinished := FALSE;
        FAbortFinished := FALSE;
        FExecutionFinished := FALSE;
        FChildrenReady := FALSE;

    E_OrchestratorTask.Execution:
        FCurrentSlot := 0;
        FHasPendingStart := FALSE;
        FExecutionFinished := FALSE;
        FResetFinished := FALSE;
        FAbortFinished := FALSE;
        IF FResult <> E_Result.Error THEN
            SelectNextSlot();
        END_IF;

    E_OrchestratorTask.Abort:
        FAbortFinished := FALSE;
END_CASE;
END_METHOD

{region 'Documentation'}
(*!
<summary>Report whether Abort remains the assigned task, including its completed phase until the task changes.</summary>
*)
{endregion}
{attribute 'monitoring' := 'call'}
PROPERTY PUBLIC IsAbortActive : BOOL //! TRUE when initialized and Abort is the assigned task, including after completion.
GET // PUBLIC
IsAbortActive := FInitialized AND (Task = E_OrchestratorTask.Abort);
END_GET
END_PROPERTY

{region 'Documentation'}
(*!
<summary>Current Abort task is finished, with reservations reconciled.</summary>
*)
{endregion}
{attribute 'monitoring' := 'call'}
PROPERTY PUBLIC IsAbortFinished : BOOL //! Current Abort task is finished, with reservations reconciled.
GET // PUBLIC
IsAbortFinished := FInitialized AND (Task = E_OrchestratorTask.Abort) AND FAbortFinished;
END_GET
END_PROPERTY

{region 'Documentation'}
(*!
<summary>Completion of the assigned task; FALSE in Idle, distinct from success.</summary>
*)
{endregion}
{attribute 'monitoring' := 'call'}
PROPERTY PUBLIC IsComplete : BOOL //! Completion of the assigned task; FALSE in Idle, distinct from success.
GET // PUBLIC
IsComplete := IsResetFinished OR IsExecutionFinished OR IsAbortFinished;
END_GET
END_PROPERTY

{region 'Documentation'}
(*!
<summary>Report whether Execution remains the assigned task, including its completed phase until the task changes.</summary>
*)
{endregion}
{attribute 'monitoring' := 'call'}
PROPERTY PUBLIC IsExecutionActive : BOOL //! TRUE when initialized and Execution is the assigned task, including after completion.
GET // PUBLIC
IsExecutionActive := FInitialized AND (Task = E_OrchestratorTask.Execution);
END_GET
END_PROPERTY

{region 'Documentation'}
(*!
<summary>Current Execution task completed all slots without a technical error.</summary>
*)
{endregion}
{attribute 'monitoring' := 'call'}
PROPERTY PUBLIC IsExecutionFinished : BOOL //! Current Execution task completed all slots without a technical error.
GET // PUBLIC
IsExecutionFinished := FInitialized AND (Task = E_OrchestratorTask.Execution) AND FExecutionFinished
    AND (FResult <> E_Result.Error);
END_GET
END_PROPERTY

{region 'Documentation'}
(*!
<summary>Report whether Initialize accepted the collection binding and cached the occupied index bounds.</summary>
*)
{endregion}
{attribute 'monitoring' := 'call'}
PROPERTY PUBLIC IsInitialized : BOOL //! Report whether Initialize accepted the collection binding and cached the occupied index bounds.
GET // PUBLIC
IsInitialized := FInitialized;
END_GET
END_PROPERTY

{region 'Documentation'}
(*!
<summary>Tests the supplied slot against the last registered child without changing state.</summary>
*)
{endregion}
METHOD PRIVATE IsLastSlot : BOOL //! TRUE when Slot is nonzero and equals the last registered child's slot in an initialized collection.
VAR_INPUT
    Slot : UINT; //! Nonzero effective execution slot to compare with the last occupied child.
END_VAR
VAR
    Child : I_Orchestratable;
END_VAR
IsLastSlot := FALSE;
IF NOT FInitialized OR (FCollection = 0) OR (Slot = 0) THEN
    RETURN;
END_IF;

Child := FCollection.GetChild(Index := FLastOccupiedIndex);
IF Child = 0 THEN
    RETURN;
END_IF;
IsLastSlot := Slot = Child.ExecutionSlot;
END_METHOD

{region 'Documentation'}
(*!
<summary>Execution may start from Idle with ready children, reconciled reservations and no held error.</summary>
*)
{endregion}
{attribute 'monitoring' := 'call'}
PROPERTY PUBLIC IsReady : BOOL //! Execution may start from Idle with ready children, reconciled reservations and no held error.
GET // PUBLIC
IsReady := FInitialized AND (Task = E_OrchestratorTask.Idle)
    AND FChildrenReady AND (FResult <> E_Result.Error);
END_GET
END_PROPERTY

{region 'Documentation'}
(*!
<summary>Report whether Reset remains the assigned task, including its completed phase until the task changes.</summary>
*)
{endregion}
{attribute 'monitoring' := 'call'}
PROPERTY PUBLIC IsResetActive : BOOL //! TRUE when initialized and Reset is the assigned task, including after completion.
GET // PUBLIC
IsResetActive := FInitialized AND (Task = E_OrchestratorTask.Reset);
END_GET
END_PROPERTY

{region 'Documentation'}
(*!
<summary>Current Reset task is finished; failed terminal children also count as finished.</summary>
*)
{endregion}
{attribute 'monitoring' := 'call'}
PROPERTY PUBLIC IsResetFinished : BOOL //! Current Reset task is finished; failed terminal children also count as finished.
GET // PUBLIC
IsResetFinished := FInitialized AND (Task = E_OrchestratorTask.Reset) AND FResetFinished;
END_GET
END_PROPERTY

{region 'Documentation'}
(*!
<summary>Checks only the selected slot for terminal completion; has no processing side effects.</summary>
*)
{endregion}
METHOD PRIVATE IsSlotCompleted : BOOL //! TRUE when every child in the selected slot is initialized and consistently Completed.
VAR
    Index : LINT;
    Child : I_Orchestratable;
END_VAR
IsSlotCompleted := FALSE;
IF (FCollection = 0) OR (FCurrentSlot = 0) THEN
    RETURN;
END_IF;
FOR Index := DINT_TO_LINT(FSlotFirstIndex) TO DINT_TO_LINT(FSlotLastIndex) DO
    Child := FCollection.GetChild(Index := LINT_TO_DINT(Index));
    IF Child = 0 THEN
        RETURN;
    END_IF;
    IF NOT Child.IsInitialized THEN
        RETURN;
    END_IF;
    IF (Child.State <> E_State.Completed) OR NOT Child.IsComplete THEN
        RETURN;
    END_IF;
END_FOR;
IsSlotCompleted := TRUE;
END_METHOD

{region 'Documentation'}
(*!
<summary>Owns pending Start confirmation, checks, cleanup and controlled child Abort.</summary>
*)
{endregion}
METHOD PRIVATE ProcessAbort
VAR
    ReservationsReleased : BOOL;
END_VAR
CheckChildStarted(ChildIndex := FPendingStartIndex,
    HasPendingStart := FHasPendingStart);
CheckChildErrors();
ReservationsReleased := FreeCompletedReservations();
UpdateReadiness();
UpdateAbortCompletion();
FChildrenReady := FChildrenReady AND ReservationsReleased;
FAbortFinished := FAbortFinished AND ReservationsReleased;
IF NOT IsAbortFinished THEN
    AbortChildren();
END_IF;
END_METHOD

{region 'Documentation'}
(*!
<summary>Owns Start confirmation, checks, reservation cleanup and slot processing.</summary>
*)
{endregion}
METHOD PRIVATE ProcessExecution
VAR
    ReservationsReleased : BOOL;
END_VAR
CheckChildStarted(ChildIndex := FPendingStartIndex,
    HasPendingStart := FHasPendingStart);
CheckChildErrors();
ReservationsReleased := FreeCompletedReservations();
UpdateReadiness();
FChildrenReady := FChildrenReady AND ReservationsReleased;
ProcessSlot();
END_METHOD

{region 'Documentation'}
(*!
<summary>Reconciles eligible reservations and readiness without dispatching child requests.</summary>
*)
{endregion}
METHOD PRIVATE ProcessIdle
VAR
    ReservationsReleased : BOOL;
END_VAR
CheckChildErrors();
ReservationsReleased := FreeCompletedReservations();
UpdateReadiness();
FChildrenReady := FChildrenReady AND ReservationsReleased;
END_METHOD

{region 'Documentation'}
(*!
<summary>Owns Reset checks, reservation cleanup, completion and capacity-bounded dispatch.</summary>
*)
{endregion}
METHOD PRIVATE ProcessReset
VAR
    ReservationsReleased : BOOL;
END_VAR
CheckChildErrors();
ReservationsReleased := FreeCompletedReservations();
UpdateReadiness();
UpdateResetCompletion();
FChildrenReady := FChildrenReady AND ReservationsReleased;
FResetFinished := FResetFinished AND ReservationsReleased;
IF NOT IsResetFinished THEN
    ResetNextChild();
END_IF;
END_METHOD

